  rq_init_comm_if_connected(9, "1")
  rq_init_comm_if_connected(2, "2")
  rq_init_comm_if_connected(3, "3")
  rq_init_comm_if_connected(4, "4")
  rq_print_connected_grippers()
  rq_gripper_communication_thread = run rq_gripper_communication()
  set_closed_norm(97.6470588235294, 1)
  set_open_norm(1.1764705882352942, 1)
  set_closed_mm(0.0, 1)
  set_open_mm(53.0, 1)
  set_closed_norm(100.0, 2)
  set_open_norm(0.0, 2)
  set_closed_mm(0.0, 2)
  set_open_mm(50.0, 2)
  set_closed_norm(100.0, 3)
  set_open_norm(0.0, 3)
  set_closed_mm(0.0, 3)
  set_open_mm(50.0, 3)
  set_closed_norm(100.0, 4)
  set_open_norm(0.0, 4)
  set_closed_mm(0.0, 4)
  set_open_mm(50.0, 4)
  rq_current_limit_enabled = False
  while(not rq_gripper_communication_thread_started):
      sync()
  end
  # end: URCap Installation Node
  # begin: URCap Installation Node
  #   Source: OPC UA, 2.0.2, Rocketfarm AS
  #   Type: OPC UA
  global opcua_daemon = rpc_factory("xmlrpc", "http://127.0.0.1:40409/RPC2")
  def opcua_client_connect(address):
  return opcua_daemon.client_connect(address)
  end
  def opcua_client_get_id(client_name):
  return opcua_daemon.client_get_id(client_name)
  end
  def opcua_client_try_connect(client_id):
  opcua_result = False
  if (opcua_daemon.client_connect(client_id)):
  sleep(0.01)
  opcua_result = opcua_daemon.client_is_connected(client_id)
  opcua_retry = 10
  while ( (not opcua_result) and (opcua_retry > 0) ):
  sleep(0.1)
  opcua_result = opcua_daemon.client_is_connected(client_id)
  opcua_retry = opcua_retry - 1
  end
  end
  return opcua_result
  end
  def opcua_client_disconnect(client_id):
  return opcua_daemon.client_disconnect(client_id)
  end
  def opcua_client_is_connected(client_id):
  return opcua_daemon.client_is_connected(client_id)
  end
  def opcua_client_read_byid(client_id, namespace_id, variable_id):
  return opcua_daemon.client_read_variable_by_id(client_id, namespace_id, variable_id)
  end
  def opcua_client_read_byname(client_id, namespace_id, variable_name):
  return opcua_daemon.client_read_variable_by_name(client_id, namespace_id, variable_name)
  end
  def opcua_client_write_byid(client_id, namespace_id, variable_id, variable_value):
  return opcua_daemon.client_write_variable_by_id(client_id, namespace_id, variable_id, variable_value)
  end
  def opcua_client_write_byname(client_id, namespace_id, variable_name, variable_value):
  return opcua_daemon.client_write_variable_by_name(client_id, namespace_id, variable_name, variable_value)
  end
  def opcua_client_last_error(client_id):
  return opcua_daemon.client_get_last_error(client_id)
  end
  def opcua_server_read_byname(variable_name):
  return opcua_daemon.server_read_variable_by_name(variable_name)
  end
  def opcua_server_write_byname(variable_name, variable_value):
  return opcua_daemon.server_write_variable_by_name(variable_name, variable_value)
  end
  def opcua_server_last_error():
  return opcua_daemon.server_get_last_error()
  end
  def opcua_error_to_string(errorCode):
  return opcua_daemon.error_code_to_string(errorCode)
  end
  # end: URCap Installation Node
  global AMR_Position=struct(position_identifier=0, x1=0, x2=0, y1=0, y2=0, theta1=0, theta2=0)
  global CAM_Pose=p[0,0,0,0,0,0]
  global CAM_Relation=""
  global CMD_Abort=  False
  global CMD_Clear=  False
  global CMD_Reset=  False
  global CMD_Start=  False
  global CMD_Suspend=  False
  global CMD_Unhold=  False
  global CMD_Unsuspend=  False
  global CNT_Rack_Output=0
  global FNC_Freedrive=  False
  global PRC_TubCounter=0
  global PRC_TubNumber=0
  global STP=0
  global easyPickCount=0
  global easyPickCount_4=0
  global easyPickCount_6=0
  global easyPickNoObj=0
  global easyPickNoObj_4=0
  global easyPickNoObj_6=0
  global easyPickParts=0
  global easyPickParts_4=0
  global easyPickParts_6=0
  global TMR_Barcode=0
  global Container_mid_1_p=p[-.379239199143, -.127191311915, .299999999998, .000000000046, -.000000000021, -1.247199999994]
  global Container_mid_1_q=[-2.477408934449926, -1.2969853503591224, -1.875639182904262, -1.539621866126728, 1.5731943360401213, -2.8009955944022717]
  global Container_capt_p=p[-.525590029047, .407247642794, .411588185841, -.000000000107, .000000000065, -2.896148821900]
  global Container_capt_q=[-3.5968351615224767, -2.0050156108707204, -0.8176271154495112, -1.8895759482008394, 1.5730967555598792, -2.2743681102957645]
  global Waypoint_67_p=p[-.400569668694, -.229578616721, .372459666505, .038872071922, .011651798558, -.774222490518]
  global Waypoint_67_q=[-2.312642001027026, -1.4746550179305746, -1.5408329553304227, -1.7283461118822494, 1.5491622513965435, -3.109828329266257]
  global Waypoint_6_p=p[.008800512419, -.547926542621, .402696567415, -.589884378425, -.007228654778, -.061268144704]
  global Waypoint_6_q=[-1.2044575850116175, -1.3416667741588135, -1.8272563219070435, -0.9884541195682068, 1.3621035814285278, -2.7712565104113978]
  global Waypoint_18_p=p[-.178371829612, -.433927395311, .368082383916, -.086593488055, .704679941724, -.007869906074]
  global Waypoint_18_q=[-1.265390698109762, -1.3355963987163086, -1.7944865226745605, -1.7402602634825648, 0.8780410885810852, -2.7713127771960657]
  global Waypoint_12_p=p[.008800512419, -.547926542621, .402696567415, -.589884378425, -.007228654778, -.061268144704]
  global Waypoint_12_q=[-1.2044575850116175, -1.3416667741588135, -1.8272563219070435, -0.9884541195682068, 1.3621035814285278, -2.7712565104113978]
  global Waypoint_19_p=p[-.178371829612, -.433927395311, .368082383916, -.086593488055, .704679941724, -.007869906074]
  global Waypoint_19_q=[-1.265390698109762, -1.3355963987163086, -1.7944865226745605, -1.7402602634825648, 0.8780410885810852, -2.7713127771960657]
  global Vial_above_p=p[.017105793010, -.652093028359, .184920586844, .000000000272, .000000000270, 1.564063451276]
  global Vial_above_q=[-1.3375440709712851, -1.9618096977868804, -1.4665759083780685, -1.2837941559171444, 1.5732503672317195, -4.47276330421513]
  global Vial_pick_point_p=p[.017105792852, -.648922724010, .093307568731, .000000000271, .000000000270, 1.564063451276]
  global Vial_pick_point_q=[-1.3366329456391917, -2.0375277831965413, -1.6071432798879028, -1.0675084332049813, 1.57309887265915, -4.471135348858068]
  global Waypoint_20_p=p[.019227646885, -.648669633640, .184920586950, .000000000000, .000000000000, .024063451426]
  global Waypoint_20_q=[-1.3331129109407733, -1.9540750545686123, -1.4775914902901128, -1.280581784992414, 1.5733500744865856, -2.928303704452631]
  global Waypoint_33_p=p[-.032361834699, -.348336136197, .391475576335, -.000008499254, .000014589902, -.004651426820]
  global Waypoint_33_q=[-1.2709335019096129, -1.1914598663441005, -1.708995335060501, -1.8117888533498316, 1.5729683532263925, -2.8379347397710237]
  global Vial_3FG_place_p=p[-.031858676359, -.349402499566, .145301120695, .000000000000, .000000000000, .000000000000]
  global Vial_3FG_place_q=[-1.2723975525801707, -1.252376585823825, -2.3128114007049496, -1.1470592278900167, 1.5730548099411423, -2.8414815174610535]
  global Waypoint_34_p=p[-.032361834699, -.348336136197, .391475576335, -.000008499254, .000014589902, -.004651426820]
  global Waypoint_34_q=[-1.2709335019096129, -1.1914598663441005, -1.708995335060501, -1.8117888533498316, 1.5729683532263925, -2.8379347397710237]
  global cap_dump_p=p[-.139168676487, -.420163541420, .146096395183, .000000000000, .000000000000, .000000000000]
  global cap_dump_q=[-1.584588644510994, -1.5093464179777323, -2.1118449369620347, -1.091059703602438, 1.5728943834877336, -3.154014906686923]
  global Waypoint_35_p=p[-.032361834699, -.348336136197, .391475576335, -.000008499254, .000014589902, -.004651426820]
  global Waypoint_35_q=[-1.2709335019096129, -1.1914598663441005, -1.708995335060501, -1.8117888533498316, 1.5729683532263925, -2.8379347397710237]
  global Waypoint_36_p=p[-.032361834699, -.348336136197, .391475576335, -.000008499254, .000014589902, -.004651426820]
  global Waypoint_36_q=[-1.2709335019096129, -1.1914598663441005, -1.708995335060501, -1.8117888533498316, 1.5729683532263925, -2.8379347397710237]
  global Waypoint_37_p=p[-.032361834699, -.348336136197, .391475576335, -.000008499254, .000014589902, -.004651426820]
  global Waypoint_37_q=[-1.2709335019096129, -1.1914598663441005, -1.708995335060501, -1.8117888533498316, 1.5729683532263925, -2.8379347397710237]
  global Vial_liq_above_p=p[-.025303660977, -.338758622354, .426628485936, -1.315858642253, .800043520260, -.928295855026]
  global Vial_liq_above_q=[-0.3789628187762659, -1.5149522957256814, -2.263045310974121, 0.7870649534412841, -0.750984017048971, -3.2237566153155726]
  global Vial_liq_pick_1_p=p[-.002660428945, -.335984893034, .159389832934, -1.150456778400, .673175527684, -1.010612657503]
  global Vial_liq_pick_1_q=[-0.3660772482501429, -1.4503649038127442, -2.4056053161621094, -1.994692941705221, 0.8039668202400208, -0.2508929411517542]
  global Vial_liq_pick_2_p=p[-.041402486291, -.356791603314, .125395323246, -1.143483969075, .651070210027, -.878721885453]
  global Vial_liq_pick_2_q=[-0.4426233705502476, -1.437252121513727, -2.551930962114307, -1.776528229806984, 0.6562026234073748, -0.43018811960029524]
  global Liquid_midway_p=p[.057575295009, -.583081747994, .306414980749, -1.351675548728, .120935756539, -.096908606303]
  global Liquid_midway_q=[-0.895174805318014, -1.7035466633238734, -2.380953073501587, 0.631549521083496, 0.7706599235534668, -2.9455552736865442]
  global shake_1_p=p[.057574880217, -.583085370269, .306422893466, -1.360996190983, -.155555042453, -.438136255921]
  global shake_1_q=[-0.8951800505267542, -1.7035466633238734, -2.380937099456787, 0.6315542894550782, 0.7706599235534669, -2.5394540616517496]
  global shake_2_p=p[.057581636113, -.583090570002, .306439684073, -1.308767904323, .368530312677, .214926493520]
  global shake_2_q=[-0.8951714674579065, -1.7035395107665003, -2.380906343460083, 0.6315504747578125, 0.7706480026245118, -3.3161255787892268]
  global drop_above_1_p=p[.268235025993, -.467784390499, .226219872376, -1.027832627524, -.430841408251, 1.004603115937]
  global drop_above_1_q=[-0.935645882283346, -1.6663371525206507, -2.4252893924713135, 0.41966931402172847, 1.8470635414123535, -3.4600217978106897]
  global drop_above_2_p=p[.219042229014, -.470775657081, .133754190740, -.313004595901, -.344395319364, 1.500564994056]
  global drop_above_2_q=[-1.0601594887284795, -1.70046459045642, -2.0799996233759863, -0.7243227230676759, 1.9429634314685202, -4.115129153870795]
  global liq_tran_1_p=p[.213067510942, -.469567035397, .100231043184, .251862243732, .217902579404, 1.592812335393]
  global liq_tran_1_q=[-0.7789645168037476, -1.822364827406652, -1.8643518410805573, -1.252158963840138, 1.3768134449520435, -3.9328333233290254]
  global Waypoint_21_p=p[.187119460405, -.493959476151, .133754190608, -.313004596540, -.344395317757, 1.500564993991]
  global Waypoint_21_q=[-1.1418328121400876, -1.7310553375189475, -2.033634768766424, -0.772026910513711, 1.958578934631971, -4.201588449364511]
  global liq_tran_2_p=p[.195957706507, -.493022614126, .100231042689, .160718757180, .109807038912, 1.525321508623]
  global liq_tran_2_q=[-0.881740380645474, -1.8244526267589851, -1.865100964490387, -1.1608866323693583, 1.4631433601076713, -3.973915130363038]
  global Vial_drop_above_p=p[.000324902251, -.648569523142, .221894115667, -.873462921366, 1.165852672573, -1.482720593185]
  global Vial_drop_above_q=[-1.0576906334721352, -2.393016994184633, -0.9236232851859159, -2.5729213042279273, 0.7903331288549689, -0.33286325848155585]
  global Vial_liq_drop_p=p[.001020867953, -.647659915585, .092915870838, -.834762611599, 1.081942994823, -1.540647900176]
  global Vial_liq_drop_q=[-1.0631954168193474, -2.4447642951220825, -1.128811017825127, -2.1983115491972294, 0.8130148661460634, -0.38984988696911316]
  global Waypoint_9_p=p[.206300564882, -.401796282405, .209941275233, .000000000049, .000000000063, 1.560839127857]
  global Waypoint_9_q=[-0.7963359454512808, -1.4686025034365713, -1.9726632321075135, -1.2709582822971974, 1.5730203818053559, -3.9272300959189193]
  global Waypoint_10_p=p[.200865824304, -.400817692024, .105072686738, .000000000049, .000000000061, 1.560839127855]
  global Waypoint_10_q=[-0.8042914374275529, -1.5824702465090397, -2.1630314773482997, -0.9667217216455377, 1.5726337265768082, -3.9342465798801403]
  global Waypoint_11_p=p[.200865824280, -.400817691999, .325177251663, .000000000049, .000000000061, 1.560839127855]
  global Waypoint_11_q=[-0.8031609769098491, -1.4190566846320642, -1.7173307870816634, -1.5758364190022327, 1.5730457436482617, -3.935202548332848]
  global Waypoint_7_p=p[-.615828862681, .233809157513, .299999999960, .005115849907, .008741794022, -2.111813105778]
  global Waypoint_7_q=[-3.2957401409809868, -1.9361965884744503, -1.2056078493731617, -1.569266158150004, 1.5650998100608482, -2.7562028470627613]
  global Waypoint_8_p=p[-.615828862366, .233809157463, .013910424379, .005115849905, .008741794020, -2.111813105780]
  global Waypoint_8_q=[-3.2964782505943173, -2.1586184138220776, -1.6500090431308791, -0.9024541777239836, 1.5648120752692236, -2.7547026290098384]
  global Waypoint_13_p=p[-.479450777041, .284140798427, .125270103493, -.276792173670, 2.098433187455, -2.121256516887]
  global Waypoint_13_q=[-2.8915050665484827, -1.9549266300597132, -2.2318272590637207, -1.6654960117735804, 0.020810842514038086, -0.4019392172442835]
  global Waypoint_70_p=p[-.472820924464, .292439826304, .207418370234, -.259787347864, -2.053484648504, 2.070709755662]
  global Waypoint_70_q=[-2.969927421603815, -2.07168115810532, -1.6835546062719366, -2.4953958198513964, 0.4489790927922641, -0.005578998612037367]
  global Waypoint_2_p=p[-.312961047461, -.152991312519, .223609826854, -.745314530454, -1.713873240489, 1.673341715282]
  global Waypoint_2_q=[-2.3560472170459192, -2.183784624139303, -1.4583134651184082, -2.6435262165465296, 1.6522362232208252, 0.043451953679323196]
  global Waypoint_3_p=p[-.113749865836, -.390110151572, .317307487562, -.519383711706, -.839884211339, 1.756868173041]
  global Waypoint_3_q=[-1.8909733931170862, -1.720626016656393, -1.5115610361099243, -2.1240560017027796, 2.1809096336364746, 0.7227501273155212]
  global Waypoint_15_p=p[.029144035010, -.436802470887, .327885032028, -.521560953301, -.623641814548, 1.862659450154]
  global Waypoint_15_q=[-1.564817253743307, -1.556895188321807, -1.6826975345611572, -1.6944714985289515, 2.2362685203552246, 1.117417335510254]
  global Waypoint_14_p=p[.068712235638, -.569419545175, .285215357659, -.679242949116, -.712065334485, 1.394044574094]
  global Waypoint_14_q=[-1.5731792953485346, -1.8029235103747094, -1.6781008808776736, -1.2218450646111982, 2.4719572998240125, 1.6394218026856375]
  global Waypoint_4_p=p[-.047220457210, -.557624911767, .136370962514, -.679242949107, -.712065334475, 1.394044574096]
  global Waypoint_4_q=[-1.7740079055958748, -2.0023561428872334, -1.7577251142892676, -1.18903287716154, 2.4487287370345143, 1.322902469273079]
  global Waypoint_25_p=p[.065436479647, -.569388431626, .287820755049, -.679242949185, -.712065334557, 1.394044574070]
  global Waypoint_25_q=[-1.5789263550890595, -1.8020194754825436, -1.6702557537748035, -1.237882536889547, 2.471995808083492, 1.6301087487321393]
  global Waypoint_39_p=p[.137772150180, -.577759956854, .299999999946, .000000000217, -.000000000207, -1.594351842625]
  global Waypoint_39_q=[-1.108978697428574, -1.776486680444405, -1.413737665315093, -1.5218908901738937, 1.5733062372356947, -1.0863866394180182]
  global Waypoint_41_p=p[.074222967010, -.565641640647, .234620140366, -.516884386806, .529223682286, -1.529619060506]
  global Waypoint_41_q=[-0.9596722604286052, -1.8767069964135548, -1.4892746174057256, -1.7813862040292285, 1.0520698599867686, -0.8199687448260349]
  global Waypoint_40_p=p[.039987741677, -.564832865048, .191055405868, -.767560686167, .343136533060, -2.241315728308]
  global Waypoint_40_q=[-1.0070649180116558, -1.8745927522477324, -1.6139175023195245, -1.6337474788493545, 1.032708081143138, -0.11587278312988403]
  global Waypoint_42_p=p[.041363380882, -.564865360786, .192805844739, .278500165520, .624117100927, .762272396553]
  global Waypoint_42_q=[-1.0050718976263102, -1.8744386685524779, -1.609151451954446, -1.6399653140247947, 1.0334006002355505, -3.254032861659603]
  global Waypoint_43_p=p[.041363380886, -.564865360780, .192805844755, .854271020883, .226833028600, 2.453002871494]
  global Waypoint_43_q=[-1.0050567614299233, -1.874341297657562, -1.6092945416026048, -1.6397580431809713, 1.0333661149462194, -5.0371728933995605]
  global Waypoint_44_p=p[.040882892233, -.564854254876, .192193763716, .110913882012, .659173708659, .275719738520]
  global Waypoint_44_q=[-1.0057704811530535, -1.8745207681598055, -1.6107765025572558, -1.637858394640876, 1.033164860873599, -2.7487836132940755]
  global Waypoint_45_p=p[.042647731639, -.564895808997, .194439423694, -.451694728506, .563172064821, -1.343350300184]
  global Waypoint_45_q=[-1.0032860829914387, -1.8741561795270565, -1.6048483308761785, -1.6453689714776623, 1.0342050634514657, -1.06078829880322]
  global Waypoint_46_p=p[.099944144487, -.566244126804, .267342790130, -.451694834765, .563172023386, -1.343350532536]
  global Waypoint_46_q=[-0.9257438092434924, -1.889970530402497, -1.3828165217629076, -1.8916791100652528, 1.0664350961373816, -0.9805910833329659]
  global Waypoint_47_p=p[.099944144444, -.566244126727, .267342790273, -.101742139519, .058679218003, -1.457888523314]
  global Waypoint_47_q=[-1.1112623176383014, -1.729989471869196, -1.5530029871033957, -1.4442770617454777, 1.4670579052775654, -1.2224020460061675]
  global Waypoint_48_p=p[-.136182767566, -.647487115908, .294247768372, -.101742139549, .058679218020, -1.457888523312]
  global Waypoint_48_q=[-1.532196177857717, -1.9115932455375173, -1.2651848069729779, -1.5055651746702665, 1.4703193777418382, -1.646379689188814]
  global Waypoint_49_p=p[-.159024328559, -.641021381179, .047691706070, -.000000000033, -.000000000027, -1.457897102937]
  global Waypoint_49_q=[-1.6098490079965062, -2.1164987141784586, -1.6156631902166785, -0.9800092198841526, 1.573231151532669, -1.722204302767242]
  global Waypoint_50_p=p[-.159024328558, -.641021381151, .291114489351, -.000000000033, -.000000000027, -1.457897102937]
  global Waypoint_50_q=[-1.609190265995684, -1.9426985888940234, -1.2189094859258596, -1.55056435122874, 1.5734384912955113, -1.7235116759964022]
  global Waypoint_53_p=p[-.050111345339, -.357608435610, .335880801283, .034180375734, .020280946727, -.284888945062]
  global Waypoint_53_q=[-1.3262308189700454, -1.2221767968893875, -1.8246061249803773, -1.7046285947349489, 1.567288986353525, -2.612420684434543]
  global Spatula_above_p=p[.246204269139, -.251090760247, .422801843345, .000124138102, -.000200585727, 3.065849606206]
  global Spatula_above_q=[-0.4045403127002336, -1.2162090781774682, -1.6111926989160175, -1.8848500617582538, 1.5728273318316153, 1.240812783494689]
  global Spatula_pick_p=p[.248137289502, -.254121766069, .229082085415, .000129501860, -.000203778890, 3.114902854826]
  global Spatula_pick_q=[-0.41237841223611227, -1.1926470264843552, -2.1253976488788204, -1.3942069101716283, 1.573236462859926, 1.185941810601359]
  global container_start_p=p[.200650292946, -.570238751958, .366326773614, 1.360500828661, .021700128770, 2.681649891414]
  global container_start_q=[-0.7669977765142582, -2.188996679669204, -0.7412727239230232, -2.581362891432544, 1.0193601740278728, 1.1884911920528847]
  global container_wp_1_p=p[.170613637794, -.572150573676, .294509026043, 1.259497117139, -.008270589399, 2.787717865625]
  global container_wp_1_q=[-0.8129253370121727, -2.0726598902108755, -1.0846040680899218, -2.2403146195823957, 1.0281191187839607, 1.0435744211830564]
  global Waypoint_55_p=p[.077280900603, -.567308602990, .212067617714, 1.259497117148, -.008270589399, 2.787717865619]
  global Waypoint_55_q=[-0.9181858327853867, -1.9744793804952083, -1.4540279077890048, -1.9155621911627945, 0.9643238328181578, 0.9457250675800015]
  global Waypoint_56_p=p[.135568164031, -.570867938153, .245215470413, 1.476861317558, -.018269607491, 2.679642659499]
  global Waypoint_56_q=[-0.8259784040282607, -2.108036981522602, -1.2111990877342924, -2.2405969375728745, 0.9451797152137279, 1.125710531287379]
  global Waypoint_74_p=p[.164827890887, -.574638012411, .193751361296, 2.053636896063, -.046507887560, 2.274278266449]
  global Waypoint_74_q=[-0.7657213433975762, -2.450387120010788, -0.9886183070290357, -2.7078095590939375, 0.8831550681477878, 1.5106229631053527]
  global Waypoint_59_p=p[.272401132286, -.578182925380, .239561357365, 2.126997331910, .113921148153, 2.155615020515]
  global Waypoint_59_q=[-0.6600120703326624, -2.700596948663229, -0.4450863301753998, -3.1158048115172328, 0.9327830672264099, 1.686402678489685]
  global Waypoint_58_p=p[.223648508176, -.578477552733, .276546452136, 2.174288010107, -.044108754041, 2.058653287678]
  global Waypoint_58_q=[-0.7290484882560344, -2.6749849159411134, -0.44426632073579775, -3.220833992584847, 0.9665895014735898, 1.686536774549042]
  global Waypoint_60_p=p[-.013316432876, -.544772031582, .383371643081, 2.208233379808, .037543335712, 2.097559881761]
  global Waypoint_60_q=[-0.9328326161883087, -2.0999933666355775, -1.1958015693111372, -3.060905141293654, 0.690378518537611, 1.7121940951337198]
  global Waypoint_61_p=p[-.412188693372, -.356446875193, .383371643081, 1.751740964455, -.739956256289, 1.600691174920]
  global Waypoint_61_q=[-1.766185342973321, -2.0999933666355775, -1.1958015693111372, -3.060905141293654, 0.690378518537611, 1.7121940951337198]
  global Waypoint_75_p=p[-.289464426518, -.270539715913, .342974028595, 1.970022309681, -.559377673198, 1.826052766187]
  global Waypoint_75_q=[-1.4144111560183354, -1.6823590986399557, -1.884837256165925, -2.819278390066456, 0.7303860451872515, 1.663813676165967]
  global After_disp_1_p=p[.234177887198, -.585611108430, .246647088243, 2.169367758708, -.046205938191, 2.085892325683]
  global After_disp_1_q=[-0.7237417555497672, -2.722180506430037, -0.41745374130672275, -3.183273654534454, 0.9607950201743994, 1.6640517363137155]
  global After_disp_2_p=p[.211085330624, -.585611108398, .185147088342, 2.169367758712, -.046205938200, 2.085892325678]
  global After_disp_2_q=[-0.7439160607523654, -2.682970768183455, -0.6530526991258174, -2.987399724069057, 0.9414795057452281, 1.665066744676871]
  global After_disp_3_p=p[.125934854156, -.585611107804, .299545938076, .959554236104, -.134386766509, 2.880651774211]
  global After_disp_3_q=[-0.9434480594885066, -2.016473586333989, -1.1036579072158617, -2.096459283015281, 1.1479556364931514, 0.8433331387406042]
  global Waypoint_62_p=p[-.542658707241, -.114281911009, .251261544113, 1.813043609523, -.679411528034, 1.655271622964]
  global Waypoint_62_q=[-2.158300033470912, -1.9418836862428677, -1.8142999147147894, -2.778920736683023, 0.21900622104017292, 1.8983390235012934]
  global Waypoint_54_p=p[-.289932145201, -.405860679656, .355713907079, 2.247669714671, -.068171894995, 2.002687374422]
  global Waypoint_54_q=[-1.3367783063113041, -1.7803423770378384, -1.77251812018054, -3.0283041649902653, 0.3777629297538141, 1.915577765236737]
  global Waypoint_63_p=p[.101294795191, -.465376052375, .381756220355, .972633305146, -.158447626639, 2.887199602585]
  global Waypoint_63_q=[-0.8528172446194038, -1.7393709485118478, -1.2544079521837954, -2.2703112963960628, 1.1965892397133469, 0.91867216443391]
  global Start_p=p[-.033064633790, -.365398531763, .389873206922, .000000000001, .000000000001, 2.725785203584]
  global Start_q=[-1.287596562866887, -1.232866726886848, -1.6880113260231102, -1.7912103151657988, 1.5729028131945846, 0.6981423183093938]
  global Waypoint_76_p=p[-.479450777041, .284140798427, .125270103493, -.276792173670, 2.098433187454, -2.121256516887]
  global Waypoint_76_q=[-2.891505066548503, -1.9549266300590151, -2.231827259067863, -1.6654960117542226, 0.020810842514162875, -0.4019392172601952]
  global TMR_Barcode_is_counting=False
  thread Timer_Thread():
    while (True):
      if (TMR_Barcode_is_counting):
        TMR_Barcode = TMR_Barcode + get_steptime()
      end
      sync()
    end
  end
  run Timer_Thread()
  def Sub_Vision_V18():
    $ 916 "Sub_Vision_V18" "noBreak"
    $ 917 "PreSettings"
    $ 918 "CAM_LM_Detected≔ False "
    global CAM_LM_Detected=  False
    $ 919 "CAM_Captures≔0"
    global CAM_Captures=0
    $ 920 "CAM_Pose≔p[0,0,0,0,0,0]"
    global CAM_Pose=p[0,0,0,0,0,0]
    $ 921 "CAM_LM_Refinmnt≔ False "
    global CAM_LM_Refinmnt=  False
    $ 922 "CAM_LM_Refined≔ False "
    global CAM_LM_Refined=  False
    $ 923 "CAM_LM_Deviatn≔p[0,0,0,0,0,0]"
    global CAM_LM_Deviatn=p[0,0,0,0,0,0]
    $ 924 "CAM_LM_ID≔0"
    global CAM_LM_ID=0
    $ 925 "CAM_Done≔ False "
    global CAM_Done=  False
    $ 926 "CAM_CNT_Obj≔0"
    global CAM_CNT_Obj=0
    $ 927 "CAM_Result = []"
    CAM_Result = []
    $ 928 "OBJ_Detected≔ False "
    global OBJ_Detected=  False
    $ 929 "FRM_Reference≔p[0,0,0,0,0,0]"
    global FRM_Reference=p[0,0,0,0,0,0]
    $ 930 "'=========='"
    # '=========='
    $ 931 "Switch Action"
    switch_1 = Action
    $ 932 "Case 13"
    if (13 == switch_1):
    elif (15 == switch_1):
      $ 1050 "Case 15"
    elif (131 == switch_1):
      $ 1096 "Case 131"
      $ 1097 "Read (SensoPart)"
      $ 1098 "Action_Info≔'search for landmark'"
      global Action_Info="search for landmark"
      $ 1099 "CAM_LM≔CAM_LMs[4]"
      global CAM_LM=CAM_LMs[4]
      $ 1100 "CAM_Relation≔CAM_LM.capture_relation"
      global CAM_Relation=CAM_LM.capture_relation
      $ 1101 "go to capture pose"
      $ 1104 "If ITM_ID≟1 and JIG≟7"
      if (ITM_ID == 1  and  JIG == 7):
        $ 1105 "PSE_T≔uLM_Cap_SSRack"
        global PSE_T=uLM_Cap_SSRack
      else:
        $ 1106 "ElseIf ITM_ID≟5 and JIG≟7"
        if (ITM_ID == 5  and  JIG == 7):
          $ 1107 "PSE_T≔FRM_Cap_SSRack"
          global PSE_T=FRM_Cap_SSRack
        else:
          $ 1108 "ElseIf ITM_ID≟13 and JIG≟7"
          if (ITM_ID == 13  and  JIG == 7):
            $ 1109 "PSE_T≔FRM_pick_rack_const"
            global PSE_T=p[-0.5568395192387274,0.34423986364170267,0.44698620470146266,-1.0069110132199915E-6,3.378712467497258E-5,-8.002029546773325E-6]
          else:
            $ 1110 "ElseIf ITM_ID≟1 and JIG≟15"
            if (ITM_ID == 1 and JIG == 15):
              $ 1111 "MoveJ"
              $ 1112 "Container_mid_1" "breakAfter"
              movej(get_inverse_kin(Container_mid_1_p, qnear=Container_mid_1_q), a=1.3962634015954636, v=1.0471975511965976, r=0.05)
              $ 1113 "Container_capt" "breakAfter"
              movej(get_inverse_kin(Container_capt_p, qnear=Container_capt_q), a=1.3962634015954636, v=1.0471975511965976)
              $ 1114 "PSE_T≔FRM_Container_S_const"
              global PSE_T=p[-0.510412665574981,0.40064363362973565,0.41159789496794374,-1.1370875604168537E-5,-3.643547521609506E-6,-2.896122366208473]
            else:
              $ 1115 "ElseIf ITM_ID≟1 and JIG≟16"
              if (ITM_ID == 1  and  JIG == 16):
                $ 1116 "MoveJ"
                $ 1117 "Waypoint_67" "breakAfter"
                movej(get_inverse_kin(Waypoint_67_p, qnear=Waypoint_67_q), a=1.3962634015954636, v=1.0471975511965976, r=0.05)
                $ 1118 "PSE_T≔FRM_Weigh_scale_const"
                global PSE_T=p[-0.5686428146306285,-0.08056859912514604,0.530011948539917,-6.439606634490112E-5,3.9349504637135406E-6,-1.5500246943089222]
              end
            end
          end
        end
      end
      $ 1119 "do_transition(PSE_T, keep_rxry=False)"
      do_transition(PSE_T, keep_rxry=False)
      $ 1120 "Set"
      set_tcp(p[0.0,0.0,0.161,3.1415,0.0,0.0])
      $ 1121 "MoveJ"
      $ 1122 "PSE_T" "breakAfter"
      movej(PSE_T, a=1.3962634015954636, v=1.7453292519943295)
      $ 1123 "CAM_Pose≔get_actual_tcp_pose()"
      global CAM_Pose= get_actual_tcp_pose ()
      $ 1124 "Loop  not CAM_Done and  not ERROR.FLAG and  not CMD_Stop"
      while (  not  CAM_Done  and    not  ERROR.FLAG  and    not  CMD_Stop):
        $ 1125 "adjust capture pose"
        $ 1126 "If CAM_LM_Detected and CAM_LM_Refinmnt"
        if (CAM_LM_Detected  and  CAM_LM_Refinmnt):
          $ 1127 "PSE_T≔p[0,0,0.300,0,0,0]"
          global PSE_T=p[0,0,0.300,0,0,0]
          $ 1128 "CAM_Pose≔PSE_T"
          global CAM_Pose=PSE_T
          $ 1129 "If  not is_reachable(FRM_Reference,[PSE_T])"
          if (  not  is_reachable(FRM_Reference,[PSE_T])):
            $ 1130 "Error"
            $ 1131 "set_error(ERROR_POSE_NOT_REACHABLE)"
            set_error(ERROR_POSE_NOT_REACHABLE)
          end
          $ 1132 "If  not ERROR.FLAG"
          if (  not  ERROR.FLAG):
            $ 1133 "MoveJ"
            $ 1134 "PSE_T" "breakAfter"
            set_tcp(p[0.0,0.0,0.161,0.0,0.0,0.0])
            movej(pose_trans(FRM_Reference, PSE_T), a=0.8726646259971648, v=1.3962634015954636)
            $ 1135 "CAM_LM_Refined≔ True "
            global CAM_LM_Refined=  True
          end
        else:
          $ 1136 "ElseIf  not CAM_LM_Detected and CAM_Captures>0"
          if (  not  CAM_LM_Detected  and  CAM_Captures>0):
            $ 1137 "MoveL"
            $ 1138 "If FRM_Reference≟p[0,0,0,0,0,0]"
            if (FRM_Reference == p[0,0,0,0,0,0]):
              $ 1139 "PSE_T≔get_random_pose(pose_ref=CAM_Pose, mode='cubic', range_max=[0.150,0.150,0.015])"
              global PSE_T=get_random_pose(pose_ref=CAM_Pose, mode="cubic", range_max=[0.150,0.150,0.015])
            else:
              $ 1144 "Else" "noBreak"
              $ 1145 "PSE_T≔get_random_pose(pose_ref=CAM_Pose, mode='rotation', range_max=[10,10,0])"
              global PSE_T=get_random_pose(pose_ref=CAM_Pose, mode="rotation", range_max=[10,10,0])
              $ 1146 "CAM_LM_Refined≔ True "
              global CAM_LM_Refined=  True
            end
            $ 1147 "If get_inverse_kin_has_solution(pose_trans(FRM_Reference, PSE_T))"
            if (get_inverse_kin_has_solution( pose_trans (FRM_Reference, PSE_T))):
              $ 1148 "Comment"
              # Comment
              $ 1149 "PSE_T" "breakAfter"
              set_tcp(p[0.0,0.0,0.161,3.1415,0.0,0.0])
              movel(pose_trans(FRM_Reference, PSE_T), a=0.03, v=0.05)
            else:
              $ 1150 "Else" "noBreak"
              $ 1151 "'If random pose is out of reach, set the initial cam pose'"
              # 'If random pose is out of reach, set the initial cam pose'
              $ 1152 "PSE_T≔CAM_Pose"
              global PSE_T=CAM_Pose
            end
          end
        end
        $ 1153 "Wait: 2.0"
        sleep(2.0)
        $ 1154 "trigger"
        $ 1155 "If ITM_ID≟1 and JIG≟7"
        if (ITM_ID == 1  and  JIG == 7):
          # begin: URCap Program Node
          #   Source: SensoPart VISOR Robotic, 2.0.0, SensoPart Industriesensorik GmbH
          #   Type: VISOR Trigger
          $ 1156 "# 1 VISOR Trigger"
          visor_changeJob(1, "Landmark_INVITE_2", 6000)
          visor_trigger(1, 6000, "arm")
          # end: URCap Program Node
        else:
          $ 1157 "ElseIf ITM_ID≟5 and JIG≟7"
          if (ITM_ID == 5  and  JIG == 7):
            # begin: URCap Program Node
            #   Source: SensoPart VISOR Robotic, 2.0.0, SensoPart Industriesensorik GmbH
            #   Type: VISOR Trigger
            $ 1158 "# 1 VISOR Trigger"
            visor_changeJob(1, "Landmark_INVITE_2", 6000)
            visor_trigger(1, 6000, "arm")
            # end: URCap Program Node
          else:
            $ 1159 "ElseIf ITM_ID≟13 and JIG≟7"
            if (ITM_ID == 13  and  JIG == 7):
              # begin: URCap Program Node
              #   Source: SensoPart VISOR Robotic, 2.0.0, SensoPart Industriesensorik GmbH
              #   Type: VISOR Trigger
              $ 1160 "# 1 VISOR Trigger"
              visor_changeJob(1, "Landmark_INVITE_2", 6000)
              visor_trigger(1, 6000, "arm")
              # end: URCap Program Node
            else:
              $ 1161 "ElseIf ITM_ID≟1 and JIG≟15"
              if (ITM_ID == 1 and JIG == 15):
                # begin: URCap Program Node
                #   Source: SensoPart VISOR Robotic, 2.0.0, SensoPart Industriesensorik GmbH
                #   Type: VISOR Trigger
                $ 1162 "# 1 VISOR Trigger"
                visor_changeJob(1, "Container", 6000)
                visor_trigger(1, 6000, "arm")
                # end: URCap Program Node
              else:
                $ 1163 "ElseIf ITM_ID≟1 and JIG≟16"
                if (ITM_ID == 1 and JIG == 16):
                  # begin: URCap Program Node
                  #   Source: SensoPart VISOR Robotic, 2.0.0, SensoPart Industriesensorik GmbH
                  #   Type: VISOR Trigger
                  $ 1164 "# 1 VISOR Trigger"
                  visor_changeJob(1, "Weigh_scale", 6000)
                  visor_trigger(1, 6000, "arm")
                  # end: URCap Program Node
                end
              end
            end
          end
        end
        $ 1168 "TM_3D_Found≔visor_partsFound(1)"
        global TM_3D_Found= visor_partsFound (1)
        $ 1169 "If TM_3D_Found>0"
        if (TM_3D_Found>0):
          $ 1170 "CAM_LM_Detected≔ True "
          global CAM_LM_Detected=  True
          $ 1171 "CAM_Captures≔0"
          global CAM_Captures=0
        else:
          $ 1172 "Else" "noBreak"
          $ 1173 "CAM_LM_Detected≔ False "
          global CAM_LM_Detected=  False
          $ 1174 "CAM_Captures≔CAM_Captures+1"
          global CAM_Captures=CAM_Captures+1
        end
        $ 1179 "result"
        $ 1180 "If CAM_LM_Detected"
        if (CAM_LM_Detected):
          $ 1181 "If (CAM_LM_Refinmnt and CAM_LM_Refined) or  not CAM_LM_Refinmnt"
          if ((CAM_LM_Refinmnt  and  CAM_LM_Refined)  or    not  CAM_LM_Refinmnt):
            $ 1239 "If ITM_ID≟1 and JIG≟7"
            if (ITM_ID == 1  and  JIG == 7):
              $ 1240 "CAM_LM_SSRack≔visor_getPose3d(1, 0)"
              global CAM_LM_SSRack= visor_getPose3d (1, 0)
            else:
              $ 1241 "ElseIf ITM_ID≟5 and JIG≟7"
              if (ITM_ID == 5  and  JIG == 7):
                $ 1242 "CAM_LM_SSRack≔visor_getPose3d(1, 0)"
                global CAM_LM_SSRack= visor_getPose3d (1, 0)
              else:
                $ 1243 "ElseIf ITM_ID≟13 and JIG≟7"
                if (ITM_ID == 13  and  JIG == 7):
                  $ 1244 "CAM_LM_Bott≔visor_getPose3d(1, 0)"
                  global CAM_LM_Bott= visor_getPose3d (1, 0)
                else:
                  $ 1245 "ElseIf ITM_ID≟1 and JIG≟15"
                  if (ITM_ID == 1 and JIG == 15):
                    $ 1246 "CAM_LM_Cont_S≔visor_getPose3d(1, 0)"
                    global CAM_LM_Cont_S= visor_getPose3d (1, 0)
                    $ 1247 "cont_img_pose≔get_actual_tcp_pose()"
                    global cont_img_pose= get_actual_tcp_pose ()
                  else:
                    $ 1248 "ElseIf ITM_ID≟1 and JIG≟16"
                    if (ITM_ID == 1 and JIG == 16):
                      $ 1249 "FRM_Weigh_scale≔visor_getPose3d(1, 0)"
                      global FRM_Weigh_scale= visor_getPose3d (1, 0)
                      $ 1250 "cont_img_pose≔get_actual_tcp_pose()"
                      global cont_img_pose= get_actual_tcp_pose ()
                    end
                  end
                end
              end
            end
            $ 1251 "CAM_Done≔ True "
            global CAM_Done=  True
          end
        else:
          $ 1252 "ElseIf  not CAM_LM_Detected and CAM_Captures<CAM_PRM_Retries"
          if (  not  CAM_LM_Detected  and  CAM_Captures<CAM_PRM_Retries):
            $ 1253 "CAM_LM_Refined≔ False "
            global CAM_LM_Refined=  False
          else:
            $ 1254 "ElseIf CAM_Captures≥CAM_PRM_Retries"
            if (CAM_Captures >= CAM_PRM_Retries):
              $ 1255 "CAM_Done≔ True "
              global CAM_Done=  True
              $ 1256 "Error"
              $ 1257 "set_error(ERROR_NO_LANDMARK)"
              set_error(ERROR_NO_LANDMARK)
            end
          end
        end
      end
    elif (151 == switch_1):
      $ 1258 "Case 151"
      $ 1259 "Detect (SensoPart)"
      $ 1260 "go to capture pose"
      $ 1261 "FRM_Reference≔FRM_Cap_SSRack"
      global FRM_Reference=FRM_Cap_SSRack
      $ 1262 "PSE_T≔p[0,0,-0.00,0,0,0]"
      global PSE_T=p[0,0,-0.00,0,0,0]
      $ 1263 "do_transition(pose_trans(FRM_Reference, PSE_T), keep_rxry=False)"
      do_transition( pose_trans (FRM_Reference, PSE_T), keep_rxry=False)
      $ 1264 "JNT_Q≔get_actual_joint_positions()"
      global JNT_Q= get_actual_joint_positions ()
      $ 1265 "JNT_Q≔[JNT_Q[0], JNT_Q[1], JNT_Q[2], JNT_Q[3], JNT_Q[4], 0]"
      global JNT_Q=[JNT_Q[0], JNT_Q[1], JNT_Q[2], JNT_Q[3], JNT_Q[4], 0]
      $ 1266 "Set"
      set_tcp(p[0.0,0.0,0.161,3.1415,0.0,0.0])
      $ 1267 "movej(get_inverse_kin(pose_trans(FRM_Reference, PSE_T), qnear=JNT_Q))"
      movej(get_inverse_kin( pose_trans (FRM_Reference, PSE_T), qnear=JNT_Q))
      $ 1268 "CAM_Pose≔pose_trans(pose_inv(FRM_Reference), get_actual_tcp_pose())"
      global CAM_Pose= pose_trans ( pose_inv (FRM_Reference),  get_actual_tcp_pose ())
      $ 1269 "Loop  not CAM_Done and  not ERROR.FLAG and  not CMD_Stop"
      while (  not  CAM_Done  and    not  ERROR.FLAG  and    not  CMD_Stop):
        $ 1270 "If  not OBJ_Detected and CAM_Captures>0"
        if (  not  OBJ_Detected  and  CAM_Captures>0):
          $ 1271 "MoveL"
          $ 1272 "If FRM_Reference≟p[0,0,0,0,0,0]"
          if (FRM_Reference == p[0,0,0,0,0,0]):
            $ 1274 "PSE_T≔get_random_pose(pose_ref=CAM_Pose, mode='rotation', range_max=[15,15,0])"
            global PSE_T=get_random_pose(pose_ref=CAM_Pose, mode="rotation", range_max=[15,15,0])
          else:
            $ 1275 "Else" "noBreak"
            $ 1276 "PSE_T≔get_random_pose(pose_ref=CAM_Pose, mode='rotation', range_max=[10,10,0])"
            global PSE_T=get_random_pose(pose_ref=CAM_Pose, mode="rotation", range_max=[10,10,0])
          end
          $ 1277 "If get_inverse_kin_has_solution(pose_trans(FRM_Reference, PSE_T))"
          if (get_inverse_kin_has_solution( pose_trans (FRM_Reference, PSE_T))):
            $ 1278 "PSE_T" "breakAfter"
            set_tcp(p[0.0,0.0,0.161,3.1415,0.0,0.0])
            movel(pose_trans(FRM_Reference, PSE_T), a=0.03, v=0.05)
          else:
            $ 1279 "Else" "noBreak"
            $ 1280 "'If random pose is out of reach, set the initial cam pose'"
            # 'If random pose is out of reach, set the initial cam pose'
            $ 1281 "PSE_T≔CAM_Pose"
            global PSE_T=CAM_Pose
            $ 1282 "PSE_T" "breakAfter"
            set_tcp(p[0.0,0.0,0.161,3.1415,0.0,0.0])
            movel(pose_trans(FRM_Reference, PSE_T), a=0.03, v=0.05)
          end
        end
        $ 1283 "Wait: 0.5"
        sleep(0.5)
        $ 1284 "Set"
        set_tcp(p[0.0,0.0,0.161,3.1415,0.0,0.0])
        # begin: URCap Program Node
        #   Source: SensoPart VISOR Robotic, 2.0.0, SensoPart Industriesensorik GmbH
        #   Type: VISOR Trigger
        $ 1285 "# 1 VISOR Trigger"
        visor_changeJob(1, "Object Detection Single", 6000)
        visor_trigger(1, 6000, "arm")
        # end: URCap Program Node
        $ 1286 "If visor_isResponseOk(1)"
        if ( visor_isResponseOk (1)):
          $ 1287 "CAM_CNT_Obj≔visor_partsFound(1)"
          global CAM_CNT_Obj= visor_partsFound (1)
          $ 1288 "CAM_OBJ_Pose≔visor_getPose3d(1, 0)"
          global CAM_OBJ_Pose= visor_getPose3d (1, 0)
          $ 1289 "If CAM_CNT_Obj>0"
          if (CAM_CNT_Obj>0):
            $ 1290 "CAM_OBJ_Color≔visor_getAdditionalData(1, 0)"
            global CAM_OBJ_Color= visor_getAdditionalData (1, 0)
            $ 1291 "CAM_DetectScore≔to_num(visor_getAdditionalData(1, 1))/1000"
            global CAM_DetectScore=to_num( visor_getAdditionalData (1, 1))/1000
            $ 1292 "OBJ_Detected≔ True "
            global OBJ_Detected=  True
          end
        else:
          $ 1293 "Else" "noBreak"
          $ 1294 "CAM_Captures≔CAM_Captures+1"
          global CAM_Captures=CAM_Captures+1
        end
        $ 1295 "If OBJ_Detected"
        if (OBJ_Detected):
          $ 1296 "Get object data"
          $ 1297 "PRC_CntDetect≔0"
          global PRC_CntDetect=0
          $ 1298 "Loop PRC_CntDetect<CAM_CNT_Obj"
          while (PRC_CntDetect<CAM_CNT_Obj):
            $ 1299 "get object and jig number"
            $ 1300 "If ITM_ID≟1 and JIG≟7"
            if (ITM_ID == 1  and  JIG == 7):
              $ 1301 "FRM_Reference≔FRM_Cap_SSRack"
              global FRM_Reference=FRM_Cap_SSRack
            else:
              $ 1302 "ElseIf ITM_ID≟5 and JIG≟7"
              if (ITM_ID == 5  and  JIG == 7):
                $ 1303 "FRM_Reference≔uLM_Cap_SSRack"
                global FRM_Reference=uLM_Cap_SSRack
              end
            end
            $ 1306 "PSE_T≔pose_trans(pose_inv(FRM_Reference), CAM_OBJ_Pose)"
            global PSE_T= pose_trans ( pose_inv (FRM_Reference), CAM_OBJ_Pose)
            $ 1307 "CAM_Result.append(get_pattern_counter(PSE_T, 'X', pattern=[10, 5], patternsize=[0.181, 0.081]))"
            CAM_Result.append(get_pattern_counter(PSE_T, "X", pattern=[10, 5], patternsize=[0.181, 0.081]))
            $ 1308 "PRC_CntDetect≔PRC_CntDetect+1"
            global PRC_CntDetect=PRC_CntDetect+1
          end
          $ 1309 "CAM_Done≔ True "
          global CAM_Done=  True
        else:
          $ 1310 "ElseIf CAM_Captures≥CAM_PRM_Retries"
          if (CAM_Captures >= CAM_PRM_Retries):
            $ 1311 "CAM_Done≔ True "
            global CAM_Done=  True
          else:
            $ 1312 "Else" "noBreak"
            $ 1313 "CAM_Captures≔CAM_Captures+1"
            global CAM_Captures=CAM_Captures+1
          end
        end
      end
    end
    $ 1314 "'=========='"
    # '=========='
    $ 1315 "PostSettings"
    $ 1316 "FRM_Reference≔p[0,0,0,0,0,0]"
    global FRM_Reference=p[0,0,0,0,0,0]
    $ 1317 "Set"
    set_tcp(p[0.0,0.0,0.161,3.1415,0.0,0.0])
    $ 1318 "CAM_Pose≔p[0,0,0,0,0,0]"
    global CAM_Pose=p[0,0,0,0,0,0]
    $ 1319 "Action≔0"
    global Action=0
    $ 1320 "Action_Info≔''"
    global Action_Info=""
  end
  def Sub_AMR_MiR_V3():
    $ 1321 "Sub_AMR_MiR_V3" "noBreak"
    $ 1322 "PreSettings"
    $ 1323 "AMR_TargetList≔[1,2,3,4,5,21,22,23,24,31,32,33,34,35,36,37,38,41]"
    global AMR_TargetList=[1,2,3,4,5,21,22,23,24,31,32,33,34,35,36,37,38,41]
    $ 1324 "AMR_Done≔ False "
    global AMR_Done=  False
    $ 1325 "AMR_PosActual≔T2O_Current_Pos"
    global AMR_PosActual=modbus_get_signal_status("T2O_Current_Pos")
    $ 1326 "AMR_Attemps≔T2O_Nav_Attemps"
    global AMR_Attemps=modbus_get_signal_status("T2O_Nav_Attemps")
    $ 1327 "AMR_Battery≔MiR_Battery_Lvl"
    global AMR_Battery=modbus_get_signal_status("MiR_Battery_Lvl")
    $ 1328 "AMR_Charging≔(T2O_Charging≟1)"
    global AMR_Charging=(modbus_get_signal_status("T2O_Charging") == 1)
    $ 1329 "AMR_Position≔struct(position_identifier=T2O_Current_Pos, x1=MiR_Position_X1, x2=MiR_Position_X2, y1=MiR_Position_Y1, y2=MiR_Position_Y2, theta1=MiR_Theta_1, theta2=MiR_Theta_2) "
    global AMR_Position=struct(position_identifier=modbus_get_signal_status("T2O_Current_Pos"), x1=modbus_get_signal_status("MiR_Position_X1"), x2=modbus_get_signal_status("MiR_Position_X2"), y1=modbus_get_signal_status("MiR_Position_Y1"), y2=modbus_get_signal_status("MiR_Position_Y2"), theta1=modbus_get_signal_status("MiR_Theta_1"), theta2=modbus_get_signal_status("MiR_Theta_2"))
    $ 1330 "If MiR_Mode≠7"
    if (modbus_get_signal_status("MiR_Mode") != 7):
      $ 1331 "Error"
      $ 1332 "set_error(ERROR_AMR_WRONG_MODE)"
      set_error(ERROR_AMR_WRONG_MODE)
      $ 1333 "AMR_Done≔ True "
      global AMR_Done=  True
    end
    $ 1334 "'=========='"
    # '=========='
    $ 1335 "Switch STATE"
    switch_1 = STATE
    $ 1336 "Case 1"
    if (1 == switch_1):
      $ 1337 "stopping"
      $ 1338 "If T2O_Done≟1 and O2T_Acknowledge≟0"
      if (modbus_get_signal_status("T2O_Done") == 1  and  modbus_get_signal_status("O2T_Acknowledge") == 0):
        $ 1339 "Set O2T_Acknowledge=1"
        modbus_set_output_register("O2T_Acknowledge", 1)
      end
      $ 1340 "Set MiR_CMD_Stop=On"
      modbus_set_output_signal("MiR_CMD_Stop", True)
      $ 1341 "AMR_Position.position_identifier = 0"
      AMR_Position.position_identifier = 0
      $ 1342 "AMR_Done≔ True "
      global AMR_Done=  True
    elif (2 == switch_1):
      $ 1343 "Case 2"
      $ 1344 "stopped"
      $ 1345 "If MiR_State≠3 and MiR_State≠5"
      if (modbus_get_signal_status("MiR_State") != 3  and  modbus_get_signal_status("MiR_State") != 5):
        $ 1346 "Set MiR_CMD_Stop=Off"
        modbus_set_output_signal("MiR_CMD_Stop", False)
      end
    elif (3 == switch_1):
      $ 1347 "Case 3"
      $ 1348 "resetting"
      $ 1349 "Set O2T_Mis_Main=Off"
      modbus_set_output_signal("O2T_Mis_Main", False)
      $ 1350 "Set O2T_Mis_Charge=Off"
      modbus_set_output_signal("O2T_Mis_Charge", False)
      $ 1351 "If MiR_Mis_Queue>0"
      if (modbus_get_signal_status("MiR_Mis_Queue")>0):
        $ 1352 "Set MiR_CMD_Clear_Q=On"
        modbus_set_output_signal("MiR_CMD_Clear_Q", True)
        $ 1353 "Wait MiR_Mis_Queue≟0"
        while (not(modbus_get_signal_status("MiR_Mis_Queue") == 0)):
          sync()
        end
        $ 1354 "Set MiR_CMD_Clear_Q=Off"
        modbus_set_output_signal("MiR_CMD_Clear_Q", False)
      end
      $ 1355 "If MiR_Error_ID≠0"
      if (modbus_get_signal_status("MiR_Error_ID") != 0):
        $ 1356 "Set MiR_CMD_Clear_E=On"
        modbus_set_output_signal("MiR_CMD_Clear_E", True)
        $ 1357 "Wait MiR_Error_ID≟0"
        while (not(modbus_get_signal_status("MiR_Error_ID") == 0)):
          sync()
        end
        $ 1358 "Set MiR_CMD_Clear_E=Off"
        modbus_set_output_signal("MiR_CMD_Clear_E", False)
      end
      $ 1359 "Set O2T_Action=0"
      modbus_set_output_register("O2T_Action", 0)
      $ 1360 "Set O2T_Acknowledge=0"
      modbus_set_output_register("O2T_Acknowledge", 0)
      $ 1361 "Set O2T_Target_Pos=0"
      modbus_set_output_register("O2T_Target_Pos", 0)
      $ 1362 "Set O2T_Footprint=0"
      modbus_set_output_register("O2T_Footprint", 0)
      $ 1363 "Set O2T_ProtectOff=0"
      modbus_set_output_register("O2T_ProtectOff", 0)
      $ 1364 "Set O2T_Dock=0"
      modbus_set_output_register("O2T_Dock", 0)
      $ 1365 "AMR_Attemps≔0"
      global AMR_Attemps=0
      $ 1366 "AMR_PosTarget≔0"
      global AMR_PosTarget=0
      $ 1367 "AMR_Step≔0"
      global AMR_Step=0
      $ 1368 "AMR_AtTarget≔ False "
      global AMR_AtTarget=  False
      $ 1369 "If MiR_State≟4 or MiR_State≟3 or MiR_State≟10"
      if (modbus_get_signal_status("MiR_State") == 4  or  modbus_get_signal_status("MiR_State") == 3  or  modbus_get_signal_status("MiR_State") == 10):
        $ 1370 "AMR_Done≔ True "
        global AMR_Done=  True
      end
    elif (5 == switch_1):
      $ 1371 "Case 5"
      $ 1372 "starting"
      $ 1373 "If MiR_State≟4"
      if (modbus_get_signal_status("MiR_State") == 4):
        $ 1374 "Set MiR_CMD_Start=On"
        modbus_set_output_signal("MiR_CMD_Start", True)
        $ 1375 "Wait MiR_State≠4"
        while (not(modbus_get_signal_status("MiR_State") != 4)):
          sync()
        end
        $ 1376 "Set MiR_CMD_Start=Off"
        modbus_set_output_signal("MiR_CMD_Start", False)
        $ 1377 "AMR_Done≔ True "
        global AMR_Done=  True
      else:
        $ 1378 "ElseIf MiR_State≟10"
        if (modbus_get_signal_status("MiR_State") == 10):
          $ 1379 "'MiR in protective stop. Wait'"
          # 'MiR in protective stop. Wait'
          $ 1380 "AMR_Done≔ True "
          global AMR_Done=  True
        else:
          $ 1381 "ElseIf MiR_State≟3"
          if (modbus_get_signal_status("MiR_State") == 3):
            $ 1382 "AMR_Done≔ True "
            global AMR_Done=  True
          end
        end
      end
    elif (6 == switch_1):
      $ 1383 "Case 6"
      $ 1384 "execute"
      $ 1385 "AMR_AtTarget≔(AMR_PosActual≟AMR_PosTarget)"
      global AMR_AtTarget=(AMR_PosActual == AMR_PosTarget)
      $ 1386 "Switch AMR_Step"
      switch_2 = AMR_Step
      $ 1387 "Case 0"
      if (0 == switch_2):
        $ 1388 "If  not AMR_AtTarget"
        if (  not  AMR_AtTarget):
          $ 1389 "AMR_Step≔1"
          global AMR_Step=1
        else:
          $ 1390 "Else" "noBreak"
          $ 1391 "AMR_Done≔ True "
          global AMR_Done=  True
        end
      elif (1 == switch_2):
        $ 1392 "Case 1"
        $ 1393 "general Settings"
        $ 1394 "Set O2T_Acknowledge=0"
        modbus_set_output_register("O2T_Acknowledge", 0)
        $ 1395 "check for error"
        $ 1396 "If OBJ_Picked and MiR_State≟10"
        if (OBJ_Picked  and  modbus_get_signal_status("MiR_State") == 10):
          $ 1397 "Error"
          $ 1398 "set_error(ERROR_ROBOT_ARM_NOT_IN_HOME_POSE)"
          set_error(ERROR_ROBOT_ARM_NOT_IN_HOME_POSE)
          $ 1399 "Action≔0"
          global Action=0
        else:
          $ 1400 "ElseIf  not found_in_list(AMR_PosTarget, AMR_TargetList)"
          if (  not  found_in_list(AMR_PosTarget, AMR_TargetList)):
            $ 1401 "Error"
            $ 1402 "set_error(ERROR_UNKNOWN_POSE)"
            set_error(ERROR_UNKNOWN_POSE)
            $ 1403 "Action≔0"
            global Action=0
          end
        end
        $ 1404 "If MiR_State≟3"
        if (modbus_get_signal_status("MiR_State") == 3):
          $ 1405 "Set MiR_CMD_Start=Off"
          modbus_set_output_signal("MiR_CMD_Start", False)
          $ 1406 "Switch Action"
          switch_3 = Action
          $ 1407 "Case 51"
          if (51 == switch_3):
            $ 1408 "Charge"
            $ 1409 "'trigger the charging mission'"
            # 'trigger the charging mission'
            $ 1410 "'target pos is predefined'"
            # 'target pos is predefined'
            $ 1411 "Set O2T_Footprint=0"
            modbus_set_output_register("O2T_Footprint", 0)
            $ 1412 "Set O2T_Action=1"
            modbus_set_output_register("O2T_Action", 1)
            $ 1413 "If MiR_Mis_Queue≟0"
            if (modbus_get_signal_status("MiR_Mis_Queue") == 0):
              $ 1414 "Set O2T_Mis_Charge=On"
              modbus_set_output_signal("O2T_Mis_Charge", True)
              $ 1415 "Wait MiR_Mis_Queue≥1"
              while (not(modbus_get_signal_status("MiR_Mis_Queue") >= 1)):
                sync()
              end
              $ 1416 "Set O2T_Mis_Charge=Off"
              modbus_set_output_signal("O2T_Mis_Charge", False)
            end
          elif (52 == switch_3):
            $ 1417 "Case 52"
            $ 1418 "Navigate"
            $ 1419 "'trigger the standard missoin'"
            # 'trigger the standard missoin'
            $ 1420 "Set O2T_Footprint=AMR_FootprintID"
            modbus_set_output_register("O2T_Footprint", AMR_FootprintID)
            $ 1421 "Set O2T_Target_Pos=AMR_PosTarget"
            modbus_set_output_register("O2T_Target_Pos", AMR_PosTarget)
            $ 1422 "Set O2T_Action=2"
            modbus_set_output_register("O2T_Action", 2)
            $ 1423 "If MiR_Mis_Queue≟0"
            if (modbus_get_signal_status("MiR_Mis_Queue") == 0):
              $ 1424 "Set O2T_Mis_Main=On"
              modbus_set_output_signal("O2T_Mis_Main", True)
              $ 1425 "Wait MiR_Mis_Queue≥1"
              while (not(modbus_get_signal_status("MiR_Mis_Queue") >= 1)):
                sync()
              end
              $ 1426 "Set O2T_Mis_Main=Off"
              modbus_set_output_signal("O2T_Mis_Main", False)
            end
          end
        else:
          $ 1427 "ElseIf MiR_State≟4"
          if (modbus_get_signal_status("MiR_State") == 4):
            $ 1428 "Set MiR_CMD_Start=On"
            modbus_set_output_signal("MiR_CMD_Start", True)
          else:
            $ 1429 "ElseIf MiR_State≟5"
            if (modbus_get_signal_status("MiR_State") == 5):
              $ 1430 "AMR_Step≔2"
              global AMR_Step=2
            else:
              $ 1431 "ElseIf MiR_State≟10"
              if (modbus_get_signal_status("MiR_State") == 10):
                $ 1432 "'AMR still in safeguard stop'"
                # 'AMR still in safeguard stop'
              end
            end
          end
        end
      elif (2 == switch_2):
        $ 1433 "Case 2"
        $ 1434 "acknowledge handshake"
        $ 1435 "If T2O_Done≟1 and O2T_Acknowledge≟0"
        if (modbus_get_signal_status("T2O_Done") == 1  and  modbus_get_signal_status("O2T_Acknowledge") == 0):
          $ 1436 "Set O2T_Acknowledge=1"
          modbus_set_output_register("O2T_Acknowledge", 1)
        else:
          $ 1437 "ElseIf T2O_Done≟0 and O2T_Acknowledge≟1"
          if (modbus_get_signal_status("T2O_Done") == 0  and  modbus_get_signal_status("O2T_Acknowledge") == 1):
            $ 1438 "Set O2T_Acknowledge=0"
            modbus_set_output_register("O2T_Acknowledge", 0)
            $ 1439 "AMR_AtTarget≔(AMR_PosActual≟AMR_PosTarget)"
            global AMR_AtTarget=(AMR_PosActual == AMR_PosTarget)
            $ 1440 "AMR_Done≔ True "
            global AMR_Done=  True
          end
        end
      end
      $ 1441 "translate errors"
      $ 1442 "If AMR_Done"
      if (AMR_Done):
        $ 1443 "Switch T2O_Error_ID"
        switch_2 = modbus_get_signal_status("T2O_Error_ID")
        $ 1444 "Case 2003"
        if (2003 == switch_2):
          $ 1445 "error"
          $ 1446 "set_error(ERROR_NOT_DOCKED)"
          set_error(ERROR_NOT_DOCKED)
        elif (2007 == switch_2):
          $ 1447 "Case 2007"
          $ 1448 "error"
          $ 1449 "set_error(ERROR_NOT_REACHABLE_TARGET)"
          set_error(ERROR_NOT_REACHABLE_TARGET)
        elif (2008 == switch_2):
          $ 1450 "Case 2008"
          $ 1451 "error"
          $ 1452 "set_error(ERROR_CHARGING_NOT_STARTED)"
          set_error(ERROR_CHARGING_NOT_STARTED)
        end
      end
    elif (7 == switch_1):
      $ 1453 "Case 7"
      $ 1454 "completing"
      $ 1455 "If MiR_Mis_Queue>0"
      if (modbus_get_signal_status("MiR_Mis_Queue")>0):
        $ 1456 "Set MiR_CMD_Abort=On"
        modbus_set_output_signal("MiR_CMD_Abort", True)
        $ 1457 "Wait MiR_Mis_Queue≟0"
        while (not(modbus_get_signal_status("MiR_Mis_Queue") == 0)):
          sync()
        end
        $ 1458 "Set MiR_CMD_Abort=Off"
        modbus_set_output_signal("MiR_CMD_Abort", False)
      end
      $ 1459 "If MiR_State≟3 or MiR_State≟10"
      if (modbus_get_signal_status("MiR_State") == 3  or  modbus_get_signal_status("MiR_State") == 10):
        $ 1460 "AMR_Done≔ True "
        global AMR_Done=  True
      end
    elif (9 == switch_1):
      $ 1461 "Case 9"
      $ 1462 "holding"
      $ 1463 "Set MiR_CMD_Abort=On"
      modbus_set_output_signal("MiR_CMD_Abort", True)
      $ 1464 "If MiR_State≟3 or MiR_State≟10"
      if (modbus_get_signal_status("MiR_State") == 3  or  modbus_get_signal_status("MiR_State") == 10):
        $ 1465 "Set MiR_CMD_Abort=Off"
        modbus_set_output_signal("MiR_CMD_Abort", False)
        $ 1466 "AMR_Done≔ True "
        global AMR_Done=  True
      end
    elif (11 == switch_1):
      $ 1467 "Case 11"
      $ 1468 "unholding"
      $ 1469 "Set MiR_CMD_Start=On"
      modbus_set_output_signal("MiR_CMD_Start", True)
      $ 1470 "If MiR_State≠4"
      if (modbus_get_signal_status("MiR_State") != 4):
        $ 1471 "Set MiR_CMD_Start=Off"
        modbus_set_output_signal("MiR_CMD_Start", False)
        $ 1472 "AMR_Step≔0"
        global AMR_Step=0
        $ 1473 "AMR_Done≔ True "
        global AMR_Done=  True
      end
    elif (12 == switch_1):
      $ 1474 "Case 12"
      $ 1475 "suspending"
      $ 1476 "'none'"
      # 'none'
    elif (14 == switch_1):
      $ 1477 "Case 14"
      $ 1478 "unsuspending"
      $ 1479 "'none'"
      # 'none'
    elif (15 == switch_1):
      $ 1480 "Case 15"
      $ 1481 "aborting"
      $ 1482 "Set MiR_CMD_Abort=On"
      modbus_set_output_signal("MiR_CMD_Abort", True)
      $ 1483 "Wait MiR_State≟3"
      while (not(modbus_get_signal_status("MiR_State") == 3)):
        sync()
      end
      $ 1484 "Set MiR_CMD_Abort=Off"
      modbus_set_output_signal("MiR_CMD_Abort", False)
    elif (17 == switch_1):
      $ 1485 "Case 17"
      $ 1486 "clearing"
      $ 1487 "If MiR_Error_ID≠0"
      if (modbus_get_signal_status("MiR_Error_ID") != 0):
        $ 1488 "Set MiR_CMD_Clear_E=On"
        modbus_set_output_signal("MiR_CMD_Clear_E", True)
        $ 1489 "Wait MiR_Error_ID≟0"
        while (not(modbus_get_signal_status("MiR_Error_ID") == 0)):
          sync()
        end
        $ 1490 "Set MiR_CMD_Clear_E=Off"
        modbus_set_output_signal("MiR_CMD_Clear_E", False)
      end
      $ 1491 "If MiR_Error_ID≟0"
      if (modbus_get_signal_status("MiR_Error_ID") == 0):
        $ 1492 "AMR_Done≔ True "
        global AMR_Done=  True
      end
    end
    $ 1493 "'=========='"
    # '=========='
    $ 1494 "PostSettings"
    $ 1495 "AMR_Position≔struct(position_identifier=T2O_Current_Pos, x1=MiR_Position_X1, x2=MiR_Position_X2, y1=MiR_Position_Y1, y2=MiR_Position_Y2, theta1=MiR_Theta_1, theta2=MiR_Theta_2) "
    global AMR_Position=struct(position_identifier=modbus_get_signal_status("T2O_Current_Pos"), x1=modbus_get_signal_status("MiR_Position_X1"), x2=modbus_get_signal_status("MiR_Position_X2"), y1=modbus_get_signal_status("MiR_Position_Y1"), y2=modbus_get_signal_status("MiR_Position_Y2"), theta1=modbus_get_signal_status("MiR_Theta_1"), theta2=modbus_get_signal_status("MiR_Theta_2"))
  end
  def Sub_Action_V4():
    $ 1496 "Sub_Action_V4" "noBreak"
    $ 1497 "PreSettings"
    $ 1498 "init poses"
    $ 1499 "PSE_A≔p[0,0,0,0,0,0]"
    global PSE_A=p[0,0,0,0,0,0]
    $ 1500 "PSE_A_H≔p[0,0,0,0,0,0]"
    global PSE_A_H=p[0,0,0,0,0,0]
    $ 1501 "PSE_T≔p[0,0,0,0,0,0]"
    global PSE_T=p[0,0,0,0,0,0]
    $ 1502 "PSE_T_H≔p[0,0,0,0,0,0]"
    global PSE_T_H=p[0,0,0,0,0,0]
    $ 1503 "PSE_G≔p[0,0,0,0,0,0]"
    global PSE_G=p[0,0,0,0,0,0]
    $ 1504 "PSE_G_H≔p[0,0,0,0,0,0]"
    global PSE_G_H=p[0,0,0,0,0,0]
    $ 1505 "PSE_R≔p[0,0,0,0,0,0]"
    global PSE_R=p[0,0,0,0,0,0]
    $ 1506 "PSE_R_H≔p[0,0,0,0,0,0]"
    global PSE_R_H=p[0,0,0,0,0,0]
    $ 1507 "JNT_Q≔[0,0,0,0,0,0]"
    global JNT_Q=[0,0,0,0,0,0]
    $ 1508 "JNT_S≔[0,0,0,0,0,0]"
    global JNT_S=[0,0,0,0,0,0]
    $ 1509 "Gripping parameters"
    $ 1510 "OBJ = find_object_by_type(OBJs, OBJ_Type)"
    OBJ = find_object_by_type(OBJs, OBJ_Type)
    $ 1511 "GRP_Open_Pos≔OBJ.dimension.diameter * 1000 + 6"
    global GRP_Open_Pos=OBJ.dimension.diameter * 1000 + 6
    $ 1512 "GRP_Offset≔OBJ.gripper_offset"
    global GRP_Offset=OBJ.gripper_offset
    $ 1513 "rq_set_force_norm(50)"
     rq_set_force_norm (50)
    $ 1514 "rq_set_speed_norm(50)"
     rq_set_speed_norm (50)
    $ 1515 "Switch ITM_ID"
    switch_1 = ITM_ID
    $ 1516 "Case 1"
    if (1 == switch_1):
      $ 1517 "uML"
      $ 1518 "JIG2 = find_object_by_type(JIGs, JIG)"
      JIG2 = find_object_by_type(JIGs, JIG)
      $ 1519 "JIG_Offset≔JIG2.jig_offset"
      global JIG_Offset=JIG2.jig_offset
      $ 1520 "Switch JIG"
      switch_2 = JIG
      $ 1521 "Case 1"
      if (1 == switch_2):
        $ 1522 "3FG"
        $ 1523 "define poses"
        $ 1524 "FRM_Reference≔ULM_3FG"
        global FRM_Reference=ULM_3FG
        $ 1525 "JNT_Q≔JNT_HOME"
        global JNT_Q=JNT_HOME
        $ 1526 "PSE_T≔pose_trans(GRP_Offset, JIG_Offset)"
        global PSE_T= pose_trans (GRP_Offset, JIG_Offset)
        $ 1527 "PSE_A≔pose_trans(PSE_T, p[0,0,0.100,0,0,0])"
        global PSE_A= pose_trans (PSE_T, p[0,0,0.100,0,0,0])
        $ 1528 "PSE_R≔pose_add(PSE_T, p[0,0,0.100,0,0,0])"
        global PSE_R= pose_add (PSE_T, p[0,0,0.100,0,0,0])
      elif (2 == switch_2):
        $ 1529 "Case 2"
        $ 1530 "Input"
        $ 1531 "'CHANGE THE REFERENCE TO THE FRAME TO MOVE IN'"
        # 'CHANGE THE REFERENCE TO THE FRAME TO MOVE IN'
        $ 1532 "define poses"
        $ 1533 "FRM_Reference≔ULM_Input"
        global FRM_Reference=ULM_Input
        $ 1534 "PSE_T≔pose_trans(pose_trans(get_pattern_pos_rectangle(OBJ_Nbr, 'X', [10,5], patternsize=[0.181,0.081]), GRP_Offset), JIG_Offset)"
        global PSE_T= pose_trans ( pose_trans (get_pattern_pos_rectangle(OBJ_Nbr, "X", [10,5], patternsize=[0.181,0.081]), GRP_Offset), JIG_Offset)
        $ 1535 "If Action≟1"
        if (Action == 1):
          $ 1536 "PSE_R≔pose_add(PSE_T, p[0,0,0.200,0,0,0])"
          global PSE_R= pose_add (PSE_T, p[0,0,0.200,0,0,0])
          $ 1537 "PSE_A≔pose_add(PSE_T, p[0,0,0.100,0,0,0])"
          global PSE_A= pose_add (PSE_T, p[0,0,0.100,0,0,0])
        else:
          $ 1538 "ElseIf Action≟2"
          if (Action == 2):
            $ 1539 "PSE_R≔pose_add(PSE_T, p[0,0,0.100,0,0,0])"
            global PSE_R= pose_add (PSE_T, p[0,0,0.100,0,0,0])
            $ 1540 "PSE_A≔pose_add(PSE_T, p[0,0,0.200,0,0,0])"
            global PSE_A= pose_add (PSE_T, p[0,0,0.200,0,0,0])
          end
        end
      elif (3 == switch_2):
        $ 1541 "Case 3"
        $ 1542 "Output"
        $ 1543 "'CHANGE THE REFERENCE TO THE FRAME TO MOVE IN'"
        # 'CHANGE THE REFERENCE TO THE FRAME TO MOVE IN'
        $ 1544 "define poses"
        $ 1545 "FRM_Reference≔ULM_Output"
        global FRM_Reference=ULM_Output
        $ 1546 "PSE_T≔pose_trans(pose_trans(get_pattern_pos_rectangle(OBJ_Nbr, 'X', [10,5], patternsize=[0.181,0.081]), GRP_Offset), JIG_Offset)"
        global PSE_T= pose_trans ( pose_trans (get_pattern_pos_rectangle(OBJ_Nbr, "X", [10,5], patternsize=[0.181,0.081]), GRP_Offset), JIG_Offset)
        $ 1548 "If Action≟1"
        if (Action == 1):
          $ 1549 "PSE_R≔pose_add(PSE_T, p[0,0,0.200,0,0,0])"
          global PSE_R= pose_add (PSE_T, p[0,0,0.200,0,0,0])
          $ 1550 "PSE_A≔pose_add(PSE_T, p[0,0,0.100,0,0,0])"
          global PSE_A= pose_add (PSE_T, p[0,0,0.100,0,0,0])
        else:
          $ 1551 "ElseIf Action≟2"
          if (Action == 2):
            $ 1552 "PSE_R≔pose_add(PSE_T, p[0,0,0.100,0,0,0])"
            global PSE_R= pose_add (PSE_T, p[0,0,0.100,0,0,0])
            $ 1553 "PSE_A≔pose_add(PSE_T, p[0,0,0.200,0,0,0])"
            global PSE_A= pose_add (PSE_T, p[0,0,0.200,0,0,0])
          end
        end
      elif (4 == switch_2):
        $ 1554 "Case 4"
        $ 1555 "jig centrifuge racks"
        $ 1556 "define poses"
        $ 1557 "FRM_Reference≔ULM_Cent_Racks"
        global FRM_Reference=ULM_Cent_Racks
        $ 1558 "PSE_T≔get_pattern_pos_rectangle(JIG_Slot, 'X', [4,1], patternsize=[0.291,0])"
        global PSE_T=get_pattern_pos_rectangle(JIG_Slot, "X", [4,1], patternsize=[0.291,0])
        $ 1559 "If OBJ_Nbr≠0"
        if (OBJ_Nbr != 0):
          $ 1560 "PSE_T≔pose_trans(pose_trans(PSE_T, get_pattern_pos_rectangle(OBJ_Nbr, 'X', [3,3], patternsize=[0.060,0.060])),p[-0.030, -0.030,0,0,0,3.927])"
          global PSE_T= pose_trans ( pose_trans (PSE_T, get_pattern_pos_rectangle(OBJ_Nbr, "X", [3,3], patternsize=[0.060,0.060])),p[-0.030, -0.030,0,0,0,3.927])
        end
        $ 1561 "PSE_T≔pose_trans(PSE_T, GRP_Offset)"
        global PSE_T= pose_trans (PSE_T, GRP_Offset)
        $ 1562 "If Action≟1"
        if (Action == 1):
          $ 1563 "PSE_R≔pose_add(PSE_T, p[0,0,0.200,0,0,0])"
          global PSE_R= pose_add (PSE_T, p[0,0,0.200,0,0,0])
          $ 1564 "PSE_A≔pose_add(PSE_T, p[0,0,0.100,0,0,0])"
          global PSE_A= pose_add (PSE_T, p[0,0,0.100,0,0,0])
        else:
          $ 1565 "ElseIf Action≟2"
          if (Action == 2):
            $ 1566 "PSE_R≔pose_add(PSE_T, p[0,0,0.100,0,0,0])"
            global PSE_R= pose_add (PSE_T, p[0,0,0.100,0,0,0])
            $ 1567 "PSE_A≔pose_add(PSE_T, p[0,0,0.200,0,0,0])"
            global PSE_A= pose_add (PSE_T, p[0,0,0.200,0,0,0])
          end
        end
      elif (6 == switch_2):
        $ 1568 "Case 6"
        $ 1569 "Caps bin"
        $ 1570 "define poses"
        $ 1571 "'Drop cap'"
        # 'Drop cap'
        $ 1572 "FRM_Reference=ULM_Cap_Bin"
        FRM_Reference=ULM_Cap_Bin
        $ 1573 "PSE_T≔pose_RPY2RotVec(p[0,0,0,0,0,0])"
        global PSE_T=pose_RPY2RotVec(p[0,0,0,0,0,0])
        $ 1574 "PSE_T_H≔pose_add(PSE_T, p[0,0,-0.011,0,0,0])"
        global PSE_T_H= pose_add (PSE_T, p[0,0,-0.011,0,0,0])
        $ 1575 "PSE_A≔pose_trans(PSE_T, p[0,0,0.1,0,0,0])"
        global PSE_A= pose_trans (PSE_T, p[0,0,0.1,0,0,0])
        $ 1576 "PSE_R_H≔pose_add(PSE_T, p[0,0,0.100,0,0,0])"
        global PSE_R_H= pose_add (PSE_T, p[0,0,0.100,0,0,0])
        $ 1577 "PSE_R≔pose_add(PSE_T, p[0,0,0.100,0,0,0])"
        global PSE_R= pose_add (PSE_T, p[0,0,0.100,0,0,0])
      elif (7 == switch_2):
        $ 1578 "Case 7"
        $ 1579 "Sarstedt"
        $ 1580 "'CHANGE THE REFERENCE TO THE FRAME TO MOVE IN'"
        # 'CHANGE THE REFERENCE TO THE FRAME TO MOVE IN'
        $ 1586 "If TASK.ID≟10"
        if (TASK.ID == 10):
          $ 1587 "Frame & Position Params"
          $ 1589 "FRM_Reference = CAM_LM_SSRack"
          FRM_Reference = CAM_LM_SSRack
          $ 1594 "PSE_T≔uLM_SS_PickPlc"
          global PSE_T=uLM_SS_PickPlc
          $ 1595 "PSE_A≔pose_trans(PSE_T, p[0,0,0.1,0,0,0])"
          global PSE_A= pose_trans (PSE_T, p[0,0,0.1,0,0,0])
          $ 1596 "PSE_R≔pose_add(PSE_T, p[0,0,0.1,0,0,0])"
          global PSE_R= pose_add (PSE_T, p[0,0,0.1,0,0,0])
        else:
          $ 1597 "ElseIf TASK.ID≟11"
          if (TASK.ID == 11):
            $ 1598 "FRM_Reference = ULM_SS_Jig"
            FRM_Reference = ULM_SS_Jig
            $ 1599 "PSE_T≔pose_RPY2RotVec(p[0,0,0,0,0,0])"
            global PSE_T=pose_RPY2RotVec(p[0,0,0,0,0,0])
            $ 1600 "PSE_T≔pose_trans(PSE_T, GRP_Offset)"
            global PSE_T=pose_trans(PSE_T, GRP_Offset)
            $ 1601 "PSE_A≔pose_trans(PSE_T, p[0,0,0.1,0,0,0])"
            global PSE_A= pose_trans (PSE_T, p[0,0,0.1,0,0,0])
            $ 1602 "PSE_R≔pose_add(PSE_T, p[0,0,0.2,0,0,0])"
            global PSE_R= pose_add (PSE_T, p[0,0,0.2,0,0,0])
          end
        end
      elif (8 == switch_2):
        $ 1603 "Case 8"
        $ 1604 "NoK"
        $ 1605 "define poses"
        $ 1606 "'NoK'"
        # 'NoK'
        $ 1607 "FRM_Reference=ULM_NoK"
        FRM_Reference=ULM_NoK
        $ 1608 "PSE_T≔pose_RPY2RotVec(p[0,0,0,0,0,0])"
        global PSE_T=pose_RPY2RotVec(p[0,0,0,0,0,0])
        $ 1609 "PSE_A≔pose_trans(PSE_T, p[0,0,0.1,0,0,0])"
        global PSE_A= pose_trans (PSE_T, p[0,0,0.1,0,0,0])
        $ 1610 "PSE_R≔pose_add(PSE_T, p[0,0,0.100,0,0,0])"
        global PSE_R= pose_add (PSE_T, p[0,0,0.100,0,0,0])
      elif (9 == switch_2):
        $ 1611 "Case 9"
        $ 1612 "Pick_bott_jig"
        $ 1613 "define poses"
        $ 1614 "'NoK'"
        # 'NoK'
        $ 1615 "FRM_Reference=ULM_bottle_pick_const"
        FRM_Reference=p[0.08175869478771049,-0.47602162643540935,0.09,0.00141829700319658,-0.0027789445191063835,0.07763675748118615]
        $ 1616 "PSE_T≔pose_RPY2RotVec(p[0,0,0,0,0,0])"
        global PSE_T=pose_RPY2RotVec(p[0,0,0,0,0,0])
        $ 1617 "PSE_A≔pose_trans(PSE_T, p[0,0,0.1,0,0,0])"
        global PSE_A= pose_trans (PSE_T, p[0,0,0.1,0,0,0])
        $ 1618 "PSE_R≔pose_add(PSE_T, p[0,0,0.100,0,0,0])"
        global PSE_R= pose_add (PSE_T, p[0,0,0.100,0,0,0])
      elif (10 == switch_2):
        $ 1619 "Case 10"
        $ 1620 "Place_bott_jig"
        $ 1621 "define poses"
        $ 1622 "'NoK'"
        # 'NoK'
        $ 1623 "FRM_Reference=ULM_bottle_plac_const"
        FRM_Reference=p[-0.09502738395762109,-0.5154087721098056,0.095,0.0014590126708889871,-0.0028280855286173575,0.07763149296298452]
        $ 1624 "PSE_T≔pose_RPY2RotVec(p[0,0,0,0,0,0])"
        global PSE_T=pose_RPY2RotVec(p[0,0,0,0,0,0])
        $ 1625 "PSE_A≔pose_trans(PSE_T, p[0,0,0.1,0,0,0])"
        global PSE_A= pose_trans (PSE_T, p[0,0,0.1,0,0,0])
        $ 1626 "PSE_R≔pose_add(PSE_T, p[0,0,0.100,0,0,0])"
        global PSE_R= pose_add (PSE_T, p[0,0,0.100,0,0,0])
      elif (11 == switch_2):
        $ 1627 "Case 11"
        $ 1628 "Place_bott_jig"
        $ 1629 "define poses"
        $ 1630 "'NoK'"
        # 'NoK'
        $ 1631 "FRM_Reference=shake"
        FRM_Reference=shake
        $ 1632 "PSE_T≔pose_RPY2RotVec(p[0,0,0,0,0,0])"
        global PSE_T=pose_RPY2RotVec(p[0,0,0,0,0,0])
        $ 1633 "PSE_A≔pose_trans(PSE_T, p[0,0,0,0,0,0])"
        global PSE_A= pose_trans (PSE_T, p[0,0,0,0,0,0])
        $ 1634 "PSE_R≔pose_add(PSE_T, p[0,0,0,0,0,0])"
        global PSE_R= pose_add (PSE_T, p[0,0,0,0,0,0])
      elif (12 == switch_2):
        $ 1635 "Case 12"
        $ 1636 "Pick_Vial_jig"
        $ 1637 "define poses"
        $ 1638 "'NoK'"
        # 'NoK'
        $ 1639 "FRM_Reference=shake"
        FRM_Reference=shake
        $ 1640 "PSE_T≔pose_RPY2RotVec(p[0,0,0,0,0,0])"
        global PSE_T=pose_RPY2RotVec(p[0,0,0,0,0,0])
        $ 1641 "PSE_A≔pose_trans(PSE_T, p[0,0,0,0,0,0])"
        global PSE_A= pose_trans (PSE_T, p[0,0,0,0,0,0])
        $ 1642 "PSE_R≔pose_add(PSE_T, p[0,0,0,0,0,0])"
        global PSE_R= pose_add (PSE_T, p[0,0,0,0,0,0])
      end
    elif (2 == switch_1):
      $ 1643 "Case 2"
      $ 1644 "Centrifuge"
      $ 1645 "'CHANGE THE REFERENCE TO THE FRAME TO MOVE IN'"
      # 'CHANGE THE REFERENCE TO THE FRAME TO MOVE IN'
      $ 1646 "define poses"
      $ 1647 "FRM_Reference≔FRM_Centrifuge"
      global FRM_Reference=FRM_Centrifuge
      $ 1648 "PSE_T≔GRP_Offset"
      global PSE_T=GRP_Offset
      $ 1649 "If Action≟8"
      if (Action == 8):
        $ 1650 "PSE_R≔pose_add(PSE_T, p[0,0,0.250,0,0,0])"
        global PSE_R= pose_add (PSE_T, p[0,0,0.250,0,0,0])
        $ 1651 "PSE_A≔pose_add(PSE_T, p[0,0,0.150,0,0,0])"
        global PSE_A= pose_add (PSE_T, p[0,0,0.150,0,0,0])
      else:
        $ 1652 "ElseIf Action≟7"
        if (Action == 7):
          $ 1653 "PSE_R≔pose_add(PSE_T, p[0,0,0.150,0,0,0])"
          global PSE_R= pose_add (PSE_T, p[0,0,0.150,0,0,0])
          $ 1654 "PSE_A≔pose_add(PSE_T, p[0,0,0.250,0,0,0])"
          global PSE_A= pose_add (PSE_T, p[0,0,0.250,0,0,0])
        end
      end
    elif (3 == switch_1):
      $ 1655 "Case 3"
      $ 1656 "Output"
      $ 1657 "'CHANGE THE REFERENCE TO THE FRAME TO MOVE IN'"
      # 'CHANGE THE REFERENCE TO THE FRAME TO MOVE IN'
      $ 1658 "define poses"
      $ 1659 "FRM_Reference≔Base_const"
      global FRM_Reference=p[0.0,0.0,0.0,0.0,0.0,0.0]
      $ 1660 "PSE_T≔p[0,0,0,0,0,0]"
      global PSE_T=p[0,0,0,0,0,0]
      $ 1661 "PSE_A≔pose_add(PSE_T, p[0,0,0.150,0,0,0])"
      global PSE_A= pose_add (PSE_T, p[0,0,0.150,0,0,0])
      $ 1662 "PSE_R≔pose_add(PSE_T, p[0,0,0.100,0,0,0])"
      global PSE_R= pose_add (PSE_T, p[0,0,0.100,0,0,0])
    elif (5 == switch_1):
      $ 1663 "Case 5"
      $ 1664 "Sarstedt Pickup Table"
      $ 1665 "'CHANGE THE REFERENCE TO THE FRAME TO MOVE IN'"
      # 'CHANGE THE REFERENCE TO THE FRAME TO MOVE IN'
      $ 1666 "Switch JIG"
      switch_2 = JIG
      $ 1667 "Case 7"
      if (7 == switch_2):
        $ 1680 "Sarstedt"
        $ 1681 "'CHANGE THE REFERENCE TO THE FRAME TO MOVE IN'"
        # 'CHANGE THE REFERENCE TO THE FRAME TO MOVE IN'
        $ 1687 "If TASK.ID≟10"
        if (TASK.ID == 10):
          $ 1688 "Frame & Position Params"
          $ 1689 "FRM_Reference = CAM_LM_SSRack"
          FRM_Reference = CAM_LM_SSRack
          $ 1690 "PSE_T≔uLM_SS_PickPlc"
          global PSE_T=uLM_SS_PickPlc
          $ 1691 "PSE_A≔pose_trans(PSE_T, p[0,0,0.1,0,0,0])"
          global PSE_A= pose_trans (PSE_T, p[0,0,0.1,0,0,0])
          $ 1692 "PSE_R≔pose_add(PSE_T, p[0,0,0.1,0,0,0])"
          global PSE_R= pose_add (PSE_T, p[0,0,0.1,0,0,0])
        end
      end
    elif (13 == switch_1):
      $ 1699 "Case 13"
      $ 1700 "Sarstedt Pickup Table"
      $ 1701 "'CHANGE THE REFERENCE TO THE FRAME TO MOVE IN'"
      # 'CHANGE THE REFERENCE TO THE FRAME TO MOVE IN'
      $ 1702 "Switch JIG"
      switch_2 = JIG
      $ 1703 "Case 7"
      if (7 == switch_2):
        $ 1716 "Bottle"
        $ 1717 "'CHANGE THE REFERENCE TO THE FRAME TO MOVE IN'"
        # 'CHANGE THE REFERENCE TO THE FRAME TO MOVE IN'
        $ 1723 "If TASK.ID≟43"
        if (TASK.ID == 43):
          $ 1724 "Frame & Position Params"
          $ 1725 "FRM_Reference = CAM_LM_Bott"
          FRM_Reference = CAM_LM_Bott
          $ 1726 "PSE_T≔uLM_SS_PickPlc"
          global PSE_T=uLM_SS_PickPlc
          $ 1727 "PSE_A≔pose_trans(PSE_T, p[0,0,0.1,0,0,0])"
          global PSE_A= pose_trans (PSE_T, p[0,0,0.1,0,0,0])
          $ 1728 "PSE_R≔pose_add(PSE_T, p[0,0,0.1,0,0,0])"
          global PSE_R= pose_add (PSE_T, p[0,0,0.1,0,0,0])
        end
      end
    end
    $ 1735 "Additional check"
    $ 1736 "If  not is_reachable(FRM_Reference,[PSE_A,PSE_A_H,PSE_T,PSE_T_H,PSE_R,PSE_R_H])"
    if (  not  is_reachable(FRM_Reference,[PSE_A,PSE_A_H,PSE_T,PSE_T_H,PSE_R,PSE_R_H])):
      $ 1737 "Error"
      $ 1738 "set_error(ERROR_POSE_NOT_REACHABLE)"
      set_error(ERROR_POSE_NOT_REACHABLE)
      $ 1739 "Action≔0"
      global Action=0
    end
    $ 1740 "'=========='"
    # '=========='
    $ 1741 "Switch Action"
    switch_1 = Action
    $ 1742 "Case 1"
    if (1 == switch_1):
      $ 1743 "Pick"
      $ 1744 "Action_Info≔'pick object'"
      global Action_Info="pick object"
      $ 1745 "do_transition(pose_trans(FRM_Reference, PSE_T), keep_rxry=OBJ_Picked)"
      do_transition( pose_trans (FRM_Reference, PSE_T), keep_rxry=OBJ_Picked)
      $ 1746 "EOAT"
      $ 1747 "If  not OBJ_Picked"
      if (  not  OBJ_Picked):
        $ 1748 "rq_move_and_wait_mm(GRP_Open_Pos)"
         rq_move_and_wait_mm (GRP_Open_Pos)
      end
      $ 1749 "If PSE_A_H≠PSE_Z"
      if (PSE_A_H != PSE_Z):
        $ 1750 "If JNT_Q≠JNT_Z"
        if (JNT_Q != JNT_Z):
          $ 1751 "movej(get_inverse_kin(pose_trans(FRM_Reference, PSE_A_H), qnear=JNT_Q), r=0.050)"
          movej(get_inverse_kin( pose_trans (FRM_Reference, PSE_A_H), qnear=JNT_Q), r=0.050)
        else:
          $ 1752 "Else" "noBreak"
          $ 1753 "movej(pose_trans(FRM_Reference, PSE_A_H), r=0.050)"
          movej( pose_trans (FRM_Reference, PSE_A_H), r=0.050)
        end
      end
      $ 1754 "If PSE_A≠PSE_Z"
      if (PSE_A != PSE_Z):
        $ 1755 "If JNT_Q≠JNT_Z"
        if (JNT_Q != JNT_Z):
          $ 1756 "movej(get_inverse_kin(pose_trans(FRM_Reference, PSE_A), qnear=JNT_Q), r=0.020)"
          movej(get_inverse_kin( pose_trans (FRM_Reference, PSE_A), qnear=JNT_Q), r=0.020)
        else:
          $ 1757 "Else" "noBreak"
          $ 1758 "movej(pose_trans(FRM_Reference, PSE_A), r=0.020)"
          movej( pose_trans (FRM_Reference, PSE_A), r=0.020)
        end
      end
      $ 1759 "MoveL"
      $ 1760 "If PSE_T_H≠PSE_Z"
      if (PSE_T_H != PSE_Z):
        $ 1761 "PSE_T_H" "breakAfter"
        movel(pose_trans(FRM_Reference, PSE_T_H), a=0.5, v=0.4, r=0.01)
      end
      $ 1762 "PSE_T" "breakAfter"
      movel(pose_trans(FRM_Reference, PSE_T), a=0.08, v=0.12)
      $ 1763 "EOAT"
      $ 1764 "rq_set_force_norm(50)"
       rq_set_force_norm (50)
      $ 1765 "rq_close_and_wait()"
       rq_close_and_wait ()
      $ 1766 "OBJ_Picked≔rq_is_object_detected()"
      global OBJ_Picked= rq_is_object_detected ()
      $ 1767 "If  not OBJ_Picked"
      if (  not  OBJ_Picked):
        $ 1768 "set_error(ERROR_NO_OBJECT_TO_PICK)"
        set_error(ERROR_NO_OBJECT_TO_PICK)
      end
      $ 1769 "EXTT"
      $ 1770 "Switch JIG"
      switch_2 = JIG
      $ 1771 "Case 1"
      if (1 == switch_2):
        $ 1772 "3FG"
        $ 1773 "If OBJ_Picked"
        if (OBJ_Picked):
          $ 1774 "Set GRP_3F_Open=On"
          set_standard_digital_out(5, True)
        end
      end
      $ 1775 "If PSE_R_H≠PSE_Z"
      if (PSE_R_H != PSE_Z):
        $ 1776 "PSE_R" "breakAfter"
        movel(pose_trans(FRM_Reference, PSE_R), a=0.5, v=0.4, r=0.01)
        $ 1777 "PSE_R_H" "breakAfter"
        movel(pose_trans(FRM_Reference, PSE_R_H), a=0.5, v=0.4)
      else:
        $ 1778 "Else" "noBreak"
        $ 1779 "PSE_R" "breakAfter"
        movel(pose_trans(FRM_Reference, PSE_R), a=0.5, v=0.4)
      end
    elif (2 == switch_1):
      $ 1780 "Case 2"
      $ 1781 "Place"
      $ 1782 "Action_Info≔'place object'"
      global Action_Info="place object"
      $ 1783 "do_transition(pose_trans(FRM_Reference, PSE_T), keep_rxry=OBJ_Picked)"
      do_transition( pose_trans (FRM_Reference, PSE_T), keep_rxry=OBJ_Picked)
      $ 1784 "EXTT"
      $ 1785 "Switch JIG"
      switch_2 = JIG
      $ 1786 "Case 1"
      if (1 == switch_2):
        $ 1787 "3FG"
        $ 1788 "If OBJ_Picked"
        if (OBJ_Picked):
          $ 1789 "Set GRP_3F_Open=On"
          set_standard_digital_out(5, True)
        end
      end
      $ 1790 "If PSE_A_H≠PSE_Z"
      if (PSE_A_H != PSE_Z):
        $ 1791 "If JNT_Q≠JNT_Z"
        if (JNT_Q != JNT_Z):
          $ 1792 "movej(get_inverse_kin(pose_trans(FRM_Reference, PSE_A_H), qnear=JNT_Q), r=0.050)"
          movej(get_inverse_kin( pose_trans (FRM_Reference, PSE_A_H), qnear=JNT_Q), r=0.050)
        else:
          $ 1793 "Else" "noBreak"
          $ 1794 "movej(pose_trans(FRM_Reference, PSE_A_H), r=0.050)"
          movej( pose_trans (FRM_Reference, PSE_A_H), r=0.050)
        end
      end
      $ 1795 "If PSE_A≠PSE_Z"
      if (PSE_A != PSE_Z):
        $ 1796 "If JNT_Q≠JNT_Z"
        if (JNT_Q != JNT_Z):
          $ 1797 "movej(get_inverse_kin(pose_trans(FRM_Reference, PSE_A), qnear=JNT_Q), r=0.020)"
          movej(get_inverse_kin( pose_trans (FRM_Reference, PSE_A), qnear=JNT_Q), r=0.020)
        else:
          $ 1798 "Else" "noBreak"
          $ 1799 "movej(pose_trans(FRM_Reference, PSE_A), r=0.020)"
          movej( pose_trans (FRM_Reference, PSE_A), r=0.020)
        end
      end
      $ 1800 "MoveL"
      $ 1801 "If PSE_T_H≠PSE_Z"
      if (PSE_T_H != PSE_Z):
        $ 1802 "PSE_T_H" "breakAfter"
        movel(pose_trans(FRM_Reference, PSE_T_H), a=0.5, v=0.4, r=0.01)
      end
      $ 1803 "PSE_T" "breakAfter"
      global move_thread_flag_1803=0
      thread move_thread_1803():
        enter_critical
        move_thread_flag_1803 = 1
        movel(pose_trans(FRM_Reference, PSE_T), a=0.05, v=0.09)
        move_thread_flag_1803 = 2
        exit_critical
      end
      move_thread_flag_1803 = 0
      move_thread_han_1803 = run move_thread_1803()
      while (True):
        local targetTcpDirection=get_target_tcp_speed()
        local stepsToRetract=tool_contact(direction=targetTcpDirection)
        if (stepsToRetract > 0):
          kill move_thread_han_1803
          stopl(0.5)
          $ 1804 "Until (tool_contact_detection)"
          break
        end
        sleep(1.0E-10)
        if (move_thread_flag_1803 > 1):
          join move_thread_han_1803
          break
        end
        sync()
      end
      $ 1805 "Force"
      sleep(0.02)
      zero_ftsensor()
      force_mode(FRM_Reference, [1, 1, 1, 0, 0, 0], [0.0, 0.0, 0.0, 0.0, 0.0, 0.0], 2, [0.1, 0.1, 0.01, 0.3490658503988659, 0.3490658503988659, 0.3490658503988659])
      $ 1806 "PSE_T" "noBreak"
      movel(pose_trans(FRM_Reference, PSE_T), a=0.04, v=0.07)
      end_force_mode()
      stopl(5.0)
      $ 1807 "EXTT"
      $ 1808 "Switch JIG"
      switch_2 = JIG
      $ 1809 "Case 1"
      if (1 == switch_2):
        $ 1810 "3FG"
        $ 1811 "If OBJ_Picked"
        if (OBJ_Picked):
          $ 1812 "Set GRP_3F_Open=Off"
          set_standard_digital_out(5, False)
          $ 1813 "Wait: 0.2"
          sleep(0.2)
        end
      end
      $ 1814 "EOAT"
      $ 1815 "rq_move_and_wait_mm(GRP_Open_Pos)"
       rq_move_and_wait_mm (GRP_Open_Pos)
      $ 1816 "OBJ_Picked≔rq_is_object_detected()"
      global OBJ_Picked= rq_is_object_detected ()
      $ 1817 "If PSE_R_H≠PSE_Z"
      if (PSE_R_H != PSE_Z):
        $ 1818 "PSE_R" "breakAfter"
        movel(pose_trans(FRM_Reference, PSE_R), a=0.5, v=0.4, r=0.01)
        $ 1819 "PSE_R_H" "breakAfter"
        movel(pose_trans(FRM_Reference, PSE_R_H), a=0.5, v=0.4)
      else:
        $ 1820 "Else" "noBreak"
        $ 1821 "PSE_R" "breakAfter"
        movel(pose_trans(FRM_Reference, PSE_R), a=0.5, v=0.4)
      end
    elif (3 == switch_1):
      $ 1822 "Case 3"
      $ 1823 "Push"
      $ 1824 "Action_Info≔'push'"
      global Action_Info="push"
    elif (4 == switch_1):
      $ 1825 "Case 4"
      $ 1826 "Pull"
      $ 1827 "Action_Info≔'pull'"
      global Action_Info="pull"
    elif (6 == switch_1):
      $ 1830 "Case 6"
      $ 1831 "Drop the cap"
      $ 1832 "If JNT_A≠[0,0,0,0,0,0]"
      if (JNT_A != [0,0,0,0,0,0]):
        $ 1833 "MoveJ"
        $ 1834 "JNT_A" "breakAfter"
        movej(JNT_A, a=1.3962634015954636, v=1.7453292519943295, r=0.02)
      else:
        $ 1835 "Else" "noBreak"
        $ 1836 "MoveJ"
        $ 1837 "PSE_A" "breakAfter"
        movej(pose_trans(FRM_Reference, PSE_A), a=1.3962634015954636, v=1.7453292519943295, r=0.02)
      end
      $ 1838 "MoveL"
      $ 1839 "PSE_T" "breakAfter"
      movel(pose_trans(FRM_Reference, PSE_T), a=0.05, v=0.09)
      $ 1840 "'ADD OPEN GRIPPER'"
      # 'ADD OPEN GRIPPER'
      # begin: URCap Program Node
      #   Source: Robotiq_Grippers, 1.8.4.4844, Robotiq Inc.
      #   Type: Gripper
      $ 1841 "Gripper Move10mm (1)"
      if not(gripper_connected[0]):
        popup("Gripper 1 must be connected to run this program.", "No connection", False, True, True)
      end
      if not(rq_is_gripper_activated("1")):
        popup("Gripper 1 is not activated. Go to Installation tab > Gripper to activate it and run the program again.", "Not activated", False, True, True)
      end
      rq_set_pos_spd_for(201, 0, 28, "1")
      rq_wait_pos_spe_for_request(201, 0, 28, "1")
      rq_go_to("1")
      rq_wait("1")
      # end: URCap Program Node
      $ 1842 "PSE_T_H" "breakAfter"
      movel(pose_trans(FRM_Reference, PSE_T_H), a=0.05, v=0.09)
      # begin: URCap Program Node
      #   Source: Robotiq_Grippers, 1.8.4.4844, Robotiq Inc.
      #   Type: Gripper
      $ 1843 "Gripper Move40mm (1)"
      if not(gripper_connected[0]):
        popup("Gripper 1 must be connected to run this program.", "No connection", False, True, True)
      end
      if not(rq_is_gripper_activated("1")):
        popup("Gripper 1 is not activated. Go to Installation tab > Gripper to activate it and run the program again.", "Not activated", False, True, True)
      end
      rq_set_pos_spd_for(63, 0, 28, "1")
      rq_wait_pos_spe_for_request(63, 0, 28, "1")
      rq_go_to("1")
      rq_wait("1")
      # end: URCap Program Node
      $ 1844 "PSE_R" "breakAfter"
      movel(pose_trans(FRM_Reference, PSE_R), a=0.5, v=0.4)
    elif (7 == switch_1):
      $ 1845 "Case 7"
      $ 1846 "Load"
      $ 1847 "Action_Info≔'load object'"
      global Action_Info="load object"
      $ 1848 "do_transition(pose_trans(FRM_Reference, PSE_T), keep_rxry=OBJ_Picked)"
      do_transition( pose_trans (FRM_Reference, PSE_T), keep_rxry=OBJ_Picked)
      $ 1849 "If PSE_A_H≠PSE_Z"
      if (PSE_A_H != PSE_Z):
        $ 1850 "If JNT_Q≠JNT_Z"
        if (JNT_Q != JNT_Z):
          $ 1851 "movej(get_inverse_kin(pose_trans(FRM_Reference, PSE_A_H), qnear=JNT_Q), r=0.050)"
          movej(get_inverse_kin( pose_trans (FRM_Reference, PSE_A_H), qnear=JNT_Q), r=0.050)
        else:
          $ 1852 "Else" "noBreak"
          $ 1853 "movej(pose_trans(FRM_Reference, PSE_A_H), r=0.050)"
          movej( pose_trans (FRM_Reference, PSE_A_H), r=0.050)
        end
      end
      $ 1854 "If PSE_A≠PSE_Z"
      if (PSE_A != PSE_Z):
        $ 1855 "If JNT_Q≠JNT_Z"
        if (JNT_Q != JNT_Z):
          $ 1856 "movej(get_inverse_kin(pose_trans(FRM_Reference, PSE_A), qnear=JNT_Q), r=0.020)"
          movej(get_inverse_kin( pose_trans (FRM_Reference, PSE_A), qnear=JNT_Q), r=0.020)
        else:
          $ 1857 "Else" "noBreak"
          $ 1858 "movej(pose_trans(FRM_Reference, PSE_A), r=0.020)"
          movej( pose_trans (FRM_Reference, PSE_A), r=0.020)
        end
      end
      $ 1859 "MoveL"
      $ 1860 "If PSE_T_H≠PSE_Z"
      if (PSE_T_H != PSE_Z):
        $ 1861 "PSE_T_H" "breakAfter"
        movel(pose_trans(FRM_Reference, PSE_T_H), a=0.5, v=0.4, r=0.01)
      end
      $ 1862 "PSE_T" "breakAfter"
      global move_thread_flag_1862=0
      thread move_thread_1862():
        enter_critical
        move_thread_flag_1862 = 1
        movel(pose_trans(FRM_Reference, PSE_T), a=0.05, v=0.09)
        move_thread_flag_1862 = 2
        exit_critical
      end
      move_thread_flag_1862 = 0
      move_thread_han_1862 = run move_thread_1862()
      while (True):
        local targetTcpDirection=get_target_tcp_speed()
        local stepsToRetract=tool_contact(direction=targetTcpDirection)
        if (stepsToRetract > 0):
          kill move_thread_han_1862
          stopl(0.5)
          $ 1863 "Until (tool_contact_detection)"
          break
        end
        sleep(1.0E-10)
        if (move_thread_flag_1862 > 1):
          join move_thread_han_1862
          break
        end
        sync()
      end
      $ 1864 "Force"
      sleep(0.02)
      zero_ftsensor()
      force_mode(FRM_Reference, [0, 1, 1, 0, 0, 1], [0.0, 0.0, 0.0, 0.0, 0.0, 0.0], 2, [0.1, 0.05, 0.02, 0.3490658503988659, 0.3490658503988659, 3.141592653589793])
      $ 1865 "PSE_T" "noBreak"
      movel(pose_trans(FRM_Reference, PSE_T), a=0.04, v=0.07)
      end_force_mode()
      stopl(5.0)
      $ 1866 "EOAT"
      $ 1867 "rq_move_and_wait_mm(GRP_Open_Pos)"
       rq_move_and_wait_mm (GRP_Open_Pos)
      $ 1868 "OBJ_Picked≔rq_is_object_detected()"
      global OBJ_Picked= rq_is_object_detected ()
      $ 1869 "If PSE_R_H≠PSE_Z"
      if (PSE_R_H != PSE_Z):
        $ 1870 "PSE_R" "breakAfter"
        movel(pose_trans(FRM_Reference, PSE_R), a=0.5, v=0.4, r=0.01)
        $ 1871 "PSE_R_H" "breakAfter"
        movel(pose_trans(FRM_Reference, PSE_R_H), a=0.5, v=0.4)
      else:
        $ 1872 "Else" "noBreak"
        $ 1873 "PSE_R" "breakAfter"
        movel(pose_trans(FRM_Reference, PSE_R), a=0.5, v=0.4)
      end
    elif (8 == switch_1):
      $ 1874 "Case 8"
      $ 1875 "Unload"
      $ 1876 "Action_Info≔'pick object'"
      global Action_Info="pick object"
      $ 1877 "do_transition(pose_trans(FRM_Reference, PSE_T), keep_rxry=OBJ_Picked)"
      do_transition( pose_trans (FRM_Reference, PSE_T), keep_rxry=OBJ_Picked)
      $ 1878 "EOAT"
      $ 1879 "If  not OBJ_Picked"
      if (  not  OBJ_Picked):
        $ 1880 "rq_move_and_wait_mm(GRP_Open_Pos)"
         rq_move_and_wait_mm (GRP_Open_Pos)
      end
      $ 1881 "If PSE_A_H≠PSE_Z"
      if (PSE_A_H != PSE_Z):
        $ 1882 "If JNT_Q≠JNT_Z"
        if (JNT_Q != JNT_Z):
          $ 1883 "movej(get_inverse_kin(pose_trans(FRM_Reference, PSE_A_H), qnear=JNT_Q), r=0.050)"
          movej(get_inverse_kin( pose_trans (FRM_Reference, PSE_A_H), qnear=JNT_Q), r=0.050)
        else:
          $ 1884 "Else" "noBreak"
          $ 1885 "movej(pose_trans(FRM_Reference, PSE_A_H), r=0.050)"
          movej( pose_trans (FRM_Reference, PSE_A_H), r=0.050)
        end
      end
      $ 1886 "If PSE_A≠PSE_Z"
      if (PSE_A != PSE_Z):
        $ 1887 "If JNT_Q≠JNT_Z"
        if (JNT_Q != JNT_Z):
          $ 1888 "movej(get_inverse_kin(pose_trans(FRM_Reference, PSE_A), qnear=JNT_Q), r=0.020)"
          movej(get_inverse_kin( pose_trans (FRM_Reference, PSE_A), qnear=JNT_Q), r=0.020)
        else:
          $ 1889 "Else" "noBreak"
          $ 1890 "movej(pose_trans(FRM_Reference, PSE_A), r=0.020)"
          movej( pose_trans (FRM_Reference, PSE_A), r=0.020)
        end
      end
      $ 1891 "MoveL"
      $ 1892 "If PSE_T_H≠PSE_Z"
      if (PSE_T_H != PSE_Z):
        $ 1893 "PSE_T_H" "breakAfter"
        movel(pose_trans(FRM_Reference, PSE_T_H), a=0.5, v=0.4, r=0.01)
      end
      $ 1894 "PSE_T" "breakAfter"
      movel(pose_trans(FRM_Reference, PSE_T), a=0.08, v=0.12)
      $ 1895 "Force"
      sleep(0.02)
      zero_ftsensor()
      force_mode(FRM_Reference, [1, 1, 0, 0, 0, 0], [0.0, 0.0, 0.0, 0.0, 0.0, 0.0], 2, [0.05, 0.05, 0.1, 0.3490658503988659, 0.3490658503988659, 0.3490658503988659])
      $ 1896 "EOAT" "noBreak"
      $ 1897 "rq_set_force_norm(50)" "noBreak"
       rq_set_force_norm (50)
      $ 1898 "rq_close_and_wait()" "noBreak"
       rq_close_and_wait ()
      $ 1899 "OBJ_Picked≔rq_is_object_detected()" "noBreak"
      global OBJ_Picked= rq_is_object_detected ()
      $ 1900 "If  not OBJ_Picked" "noBreak"
      if (  not  OBJ_Picked):
        $ 1901 "set_error(ERROR_NO_OBJECT_TO_PICK)" "noBreak"
        set_error(ERROR_NO_OBJECT_TO_PICK)
      end
      $ 1902 "If PSE_R_H≠PSE_Z" "noBreak"
      if (PSE_R_H != PSE_Z):
        $ 1903 "PSE_R" "noBreak"
        movel(pose_trans(FRM_Reference, PSE_R), a=0.5, v=0.4, r=0.01)
        $ 1904 "PSE_R_H" "noBreak"
        movel(pose_trans(FRM_Reference, PSE_R_H), a=0.5, v=0.4)
      else:
        $ 1905 "Else" "noBreak"
        $ 1906 "PSE_R" "noBreak"
        movel(pose_trans(FRM_Reference, PSE_R), a=0.5, v=0.4)
      end
      end_force_mode()
      stopl(5.0)
    elif (11 == switch_1):
      $ 1907 "Case 11"
      $ 1908 "Place without opening gripper"
      $ 1909 "Action_Info≔'place object without gripper opening'"
      global Action_Info="place object without gripper opening"
      $ 1911 "movel(FRM_Container_S, a=0.025, v=0.015, r=0.00001)"
      movel(FRM_Container_S, a=0.025, v=0.015, r=0.00001)
      $ 1912 "EXTT"
      $ 1913 "Switch JIG"
      switch_2 = JIG
      $ 1914 "Case 1"
      if (1 == switch_2):
        $ 1915 "3FG"
        $ 1916 "If OBJ_Picked"
        if (OBJ_Picked):
          $ 1917 "Set GRP_3F_Open=On"
          set_standard_digital_out(5, True)
        end
      end
      $ 1918 "If PSE_A_H≠PSE_Z"
      if (PSE_A_H != PSE_Z):
        $ 1919 "If JNT_Q≠JNT_Z"
        if (JNT_Q != JNT_Z):
          $ 1920 "movej(get_inverse_kin(pose_trans(FRM_Reference, PSE_A_H), qnear=JNT_Q), r=0.050)"
          movej(get_inverse_kin( pose_trans (FRM_Reference, PSE_A_H), qnear=JNT_Q), r=0.050)
        else:
          $ 1921 "Else" "noBreak"
          $ 1922 "movej(pose_trans(FRM_Reference, PSE_A_H), r=0.050)"
          movej( pose_trans (FRM_Reference, PSE_A_H), r=0.050)
        end
      end
      $ 1923 "If PSE_A≠PSE_Z"
      if (PSE_A != PSE_Z):
        $ 1924 "If JNT_Q≠JNT_Z"
        if (JNT_Q != JNT_Z):
          $ 1925 "movej(get_inverse_kin(pose_trans(FRM_Reference, PSE_A), qnear=JNT_Q), r=0.020)"
          movej(get_inverse_kin( pose_trans (FRM_Reference, PSE_A), qnear=JNT_Q), r=0.020)
        else:
          $ 1926 "Else" "noBreak"
          $ 1927 "movej(pose_trans(FRM_Reference, PSE_A), r=0.020)"
          movej( pose_trans (FRM_Reference, PSE_A), r=0.020)
        end
      end
      $ 1928 "MoveL"
      $ 1929 "If PSE_T_H≠PSE_Z"
      if (PSE_T_H != PSE_Z):
        $ 1930 "PSE_T_H" "breakAfter"
        movel(pose_trans(FRM_Reference, PSE_T_H), a=0.5, v=0.4, r=0.01)
      end
      $ 1931 "PSE_T" "breakAfter"
      global move_thread_flag_1931=0
      thread move_thread_1931():
        enter_critical
        move_thread_flag_1931 = 1
        movel(pose_trans(FRM_Reference, PSE_T), a=0.05, v=0.09)
        move_thread_flag_1931 = 2
        exit_critical
      end
      move_thread_flag_1931 = 0
      move_thread_han_1931 = run move_thread_1931()
      while (True):
        local targetTcpDirection=get_target_tcp_speed()
        local stepsToRetract=tool_contact(direction=targetTcpDirection)
        if (stepsToRetract > 0):
          kill move_thread_han_1931
          stopl(0.5)
          $ 1932 "Until (tool_contact_detection)"
          break
        end
        sleep(1.0E-10)
        if (move_thread_flag_1931 > 1):
          join move_thread_han_1931
          break
        end
        sync()
      end
      $ 1933 "Force"
      sleep(0.02)
      zero_ftsensor()
      force_mode(FRM_Reference, [1, 1, 1, 0, 0, 0], [0.0, 0.0, 0.0, 0.0, 0.0, 0.0], 2, [0.1, 0.1, 0.01, 0.3490658503988659, 0.3490658503988659, 0.3490658503988659])
      $ 1934 "PSE_T" "noBreak"
      movel(pose_trans(FRM_Reference, PSE_T), a=0.04, v=0.07)
      end_force_mode()
      stopl(5.0)
      $ 1935 "EXTT"
      $ 1936 "Switch JIG"
      switch_2 = JIG
      $ 1937 "Case 1"
      if (1 == switch_2):
        $ 1938 "3FG"
        $ 1939 "If OBJ_Picked"
        if (OBJ_Picked):
          $ 1940 "Set GRP_3F_Open=Off"
          set_standard_digital_out(5, False)
          $ 1941 "Wait: 0.2"
          sleep(0.2)
        end
      end
      $ 1942 "EOAT"
      $ 1943 "Comment"
      # Comment
    elif (12 == switch_1):
      $ 1944 "Case 12"
      $ 1945 "Decap"
      $ 1946 "Action_Info≔'decapping'"
      global Action_Info="decapping"
      $ 1947 "Set GRP_3F_Enable=On"
      set_standard_digital_out(4, True)
      $ 1948 "Set GRP_3F_Decap=On"
      set_standard_digital_out(3, True)
      $ 1949 "Force"
      sleep(0.02)
      zero_ftsensor()
      force_mode(tool_pose(), [0, 0, 1, 0, 0, 0], [0.0, 0.0, 5.0, 0.0, 0.0, 0.0], 2, [0.1, 0.1, 0.15, 0.3490658503988659, 0.3490658503988659, 0.3490658503988659])
      $ 1950 "check_decapping(offset=0.015, timeout=5, abort=CMD_Hold)" "noBreak"
      check_decapping(offset=0.015, timeout=5, abort=CMD_Hold)
      end_force_mode()
      stopl(5.0)
      $ 1951 "Set GRP_3F_Decap=Off"
      set_standard_digital_out(3, False)
      $ 1952 "Set GRP_3F_Enable=Off"
      set_standard_digital_out(4, False)
      $ 1953 "MoveL"
      $ 1954 "PSE_R" "breakAfter"
      movel(pose_trans(FRM_Reference, PSE_R), a=0.8, v=0.15)
    elif (13 == switch_1):
      $ 1955 "Case 13"
      $ 1956 "TMR_Barcode: Reset"
      TMR_Barcode = 0
      $ 1957 "Read"
      $ 1958 "TMR_Barcode: Start"
      TMR_Barcode_is_counting = True
      $ 1959 "If TMR_Barcode<PRM_TO_Read_BC"
      global thread_flag_1959=0
      thread Thread_if_1959():
        $ 1960 "KeyenceTrigger"
        $ 1961 "Set OClearResult=HI:Pulse 0.2"
        thread SinglePulse42():
          write_output_boolean_register(2, True)
          sleep(0.2)
          write_output_boolean_register(2, False)
        end
        singlePulse42 = run SinglePulse42()
        $ 1962 "Wait: 0.5"
        sleep(0.5)
        $ 1963 "Set OTriggerBarcode=Off"
        write_output_boolean_register(1, False)
        $ 1964 "Wait: 0.5"
        sleep(0.5)
        $ 1965 "Set OTriggerBarcode=On"
        write_output_boolean_register(1, True)
        $ 1966 "Wait: 0.5"
        sleep(0.5)
        $ 1967 "Preorient"
        $ 1968 "TMR_Barcode: Reset"
        TMR_Barcode = 0
        $ 1969 "If ICmdExctd"
        if (read_input_boolean_register(12)):
          $ 1970 "Set GRP_3F_Decap=On"
          set_standard_digital_out(3, True)
          $ 1971 "Set GRP_3F_Enable=On"
          set_standard_digital_out(4, True)
          $ 1972 "Loop ICmdExctd"
          while (read_input_boolean_register(12)):
            $ 1973 "KeyenceTrigger"
            $ 1974 "Set OClearResult=HI:Pulse 0.1"
            thread SinglePulse43():
              write_output_boolean_register(2, True)
              sleep(0.1)
              write_output_boolean_register(2, False)
            end
            singlePulse43 = run SinglePulse43()
            $ 1975 "Wait: 0.3"
            sleep(0.3)
            $ 1976 "Set OTriggerBarcode=Off"
            write_output_boolean_register(1, False)
            $ 1977 "Wait: 0.3"
            sleep(0.3)
            $ 1978 "Set OTriggerBarcode=On"
            write_output_boolean_register(1, True)
            $ 1979 "Wait: 0.1"
            sleep(0.1)
          end
        end
        $ 1980 "If  not ICmdExctd"
        if (  not  read_input_boolean_register(12)):
          $ 1981 "Set GRP_3F_Decap=On"
          set_standard_digital_out(3, True)
          $ 1982 "Set GRP_3F_Enable=On"
          set_standard_digital_out(4, True)
          $ 1983 "Wait ICmdExctd=HI"
          while (read_input_boolean_register(12) == False):
            sync()
          end
        end
        $ 1984 "Set GRP_3F_Decap=Off"
        set_standard_digital_out(3, False)
        $ 1985 "Set GRP_3F_Enable=Off"
        set_standard_digital_out(4, False)
        $ 1986 "OBJ_Brc_OK≔ True "
        global OBJ_Brc_OK=  True
        thread_flag_1959 = 1
      end
      if (TMR_Barcode<PRM_TO_Read_BC):
        global thread_handler_1959=run Thread_if_1959()
        while (thread_flag_1959 == 0):
          if not(TMR_Barcode<PRM_TO_Read_BC):
            kill thread_handler_1959
            thread_flag_1959 = 2
          else:
            sync()
          end
        end
      else:
        thread_flag_1959 = 2
      end
      if (thread_flag_1959 == 2):
        $ 1987 "Else" "noBreak"
        $ 1988 "exeption"
        $ 1989 "error"
        $ 1991 "OBJ_Brc_OK≔ False "
        global OBJ_Brc_OK=  False
      end
      $ 1992 "Set GRP_3F_Decap=Off"
      set_standard_digital_out(3, False)
      $ 1993 "Set GRP_3F_Enable=Off"
      set_standard_digital_out(4, False)
      $ 1994 "Set OTriggerBarcode=Off"
      write_output_boolean_register(1, False)
    elif (15 == switch_1):
      $ 1995 "Case 15"
      $ 1996 "Detect"
      $ 1997 "Action_Info≔'detect'"
      global Action_Info="detect"
    elif (30 == switch_1):
      $ 1998 "Case 30"
      $ 1999 "Shake"
      $ 2000 "Action_Info≔'shake'"
      global Action_Info="shake"
      $ 2001 "do_transition(pose_trans(FRM_Reference, PSE_T), keep_rxry=OBJ_Picked)"
      do_transition( pose_trans (FRM_Reference, PSE_T), keep_rxry=OBJ_Picked)
      $ 2002 "If PSE_A_H≠PSE_Z"
      if (PSE_A_H != PSE_Z):
        $ 2003 "If JNT_Q≠JNT_Z"
        if (JNT_Q != JNT_Z):
          $ 2004 "movej(get_inverse_kin(pose_trans(FRM_Reference, PSE_A_H), qnear=JNT_Q), r=0.050)"
          movej(get_inverse_kin( pose_trans (FRM_Reference, PSE_A_H), qnear=JNT_Q), r=0.050)
        else:
          $ 2005 "Else" "noBreak"
          $ 2006 "movej(pose_trans(FRM_Reference, PSE_A_H), r=0.050)"
          movej( pose_trans (FRM_Reference, PSE_A_H), r=0.050)
        end
      end
      $ 2007 "If PSE_A≠PSE_Z"
      if (PSE_A != PSE_Z):
        $ 2008 "If JNT_Q≠JNT_Z"
        if (JNT_Q != JNT_Z):
          $ 2009 "movej(get_inverse_kin(pose_trans(FRM_Reference, PSE_A), qnear=JNT_Q), r=0.020)"
          movej(get_inverse_kin( pose_trans (FRM_Reference, PSE_A), qnear=JNT_Q), r=0.020)
        else:
          $ 2010 "Else" "noBreak"
          $ 2011 "movej(pose_trans(FRM_Reference, PSE_A), r=0.020)"
          movej( pose_trans (FRM_Reference, PSE_A), r=0.020)
        end
      end
      $ 2012 "MoveL"
      $ 2013 "If PSE_T_H≠PSE_Z"
      if (PSE_T_H != PSE_Z):
        $ 2014 "PSE_T_H" "breakAfter"
        movel(pose_trans(FRM_Reference, PSE_T_H), a=0.5, v=0.4, r=0.01)
      end
      $ 2015 "PSE_T" "breakAfter"
      movel(pose_trans(FRM_Reference, PSE_T), a=0.08, v=0.12)
      $ 2016 "EXTT"
      $ 2017 "Comment"
      # Comment
      $ 2018 "MoveJ"
      $ 2019 "Waypoint_6" "breakAfter"
      movej(get_inverse_kin(Waypoint_6_p, qnear=Waypoint_6_q), a=1.3962634015954636, v=1.0471975511965976)
      $ 2020 "MoveJ"
      $ 2021 "Waypoint_18" "breakAfter"
      movej(get_inverse_kin(Waypoint_18_p, qnear=Waypoint_18_q), a=1.3962634015954636, v=1.0471975511965976)
      $ 2022 "MoveJ"
      $ 2023 "Waypoint_12" "breakAfter"
      movej(get_inverse_kin(Waypoint_12_p, qnear=Waypoint_12_q), a=1.3962634015954636, v=1.0471975511965976)
      $ 2024 "MoveJ"
      $ 2025 "Waypoint_19" "breakAfter"
      movej(get_inverse_kin(Waypoint_19_p, qnear=Waypoint_19_q), a=1.3962634015954636, v=1.0471975511965976)
      $ 2026 "If PSE_R_H≠PSE_Z"
      if (PSE_R_H != PSE_Z):
        $ 2027 "PSE_R" "breakAfter"
        movel(pose_trans(FRM_Reference, PSE_R), a=0.5, v=0.4, r=0.01)
        $ 2028 "PSE_R_H" "breakAfter"
        movel(pose_trans(FRM_Reference, PSE_R_H), a=0.5, v=0.4)
      else:
        $ 2029 "Else" "noBreak"
        $ 2030 "PSE_R" "breakAfter"
        movel(pose_trans(FRM_Reference, PSE_R), a=0.5, v=0.4)
      end
    elif (31 == switch_1):
      $ 2031 "Case 31"
